// TIA Portal project "ağırlık" (V16)
// Vorlageprojekt für das Buch mit Zielsystem S7-1200

(* hardware
DEVICE "S7-1200-Station_1"  S7-1200 Station
   slot 0: "Baugruppenträger_0"  Rack  V1.0
   slot 1: "PLC_1"  CPU 1211C DC/DC/DC  6ES7 211-1AE40-0XB0  V4.1
DEVICE "HMI_1"  KTP700 Basic PN
   slot 0: "HMI_1"  KTP700 Basic PN  6AV2 123-2GB03-0AX0  16.0.0.0
   slot 1: "HMI_RT_1"  KTP700 Basic PN  6AV2 123-2GB03-0AX0  16.0.0.0
   slot 5: "HMI_1.IE_CP_1"  PROFINET Interface  16.0.0.0
      slot 1: "PROFINET Interface_1"  PROFINET Interface
         slot 1: "Port_1"  Port
*)

// ===== PLC "PLC_1"  CPU 1211C DC/DC/DC =====

VAR_GLOBAL   // PLC tag table "Default Table"
   "At scale entry" AT %I0.0 : Bool;
   "At scale" AT %I0.1 : Bool;
   "At scale exit" AT %I0.2 : Bool;
   "Left Pallet Sensor" AT %I0.3 : Bool;
   "At exit left" AT %I0.4 : Bool;
   "Front Palet sensor" AT %I0.5 : Bool;
   "At exit front" AT %I0.6 : Bool;
   "Right Pallet Sensor" AT %I0.7 : Bool;
   "At exit right" AT %I1.0 : Bool;
   "Start" AT %I1.1 : Bool;
   "Reset" AT %I1.2 : Bool;
   "Stop" AT %I1.3 : Bool;
   "FACTORY I/O (Running)" AT %I1.5 : Bool;
   "Pick & Place 1 (Box Detected)" AT %I1.6 : Bool;
   "Pick & Place 2 (Box Detected)" AT %I1.7 : Bool;
   "Pick & Place 3 (Box Detected)" AT %I2.0 : Bool;
   "Entry conveyor" AT %Q0.0 : Bool;
   "Load scale" AT %Q0.1 : Bool;
   "Send left" AT %Q0.2 : Bool;
   "Left conveyor" AT %Q0.3 : Bool;
   "Send right" AT %Q0.4 : Bool;
   "Right conveyor" AT %Q0.5 : Bool;
   "Send forward" AT %Q0.6 : Bool;
   "Front conveyor" AT %Q0.7 : Bool;
   "Start light" AT %Q1.0 : Bool;
   "Reset light" AT %Q1.1 : Bool;
   "Stop light" AT %Q1.2 : Bool;
   "Left Roller conveyor" AT %Q1.3 : Bool;
   "Right Roller Conveyor" AT %Q1.4 : Bool;
   "Front Roller conveyor" AT %Q1.5 : Bool;
END_VAR

VAR_GLOBAL   // PLC tag table "Tag table_1"
   "Pick & Place 1 X Position (V)" AT %ID34 : Real;
   "Pick & Place 1 Z Position (V)" AT %ID38 : Real;
   "Pick & Place 2 X Position (V)" AT %ID42 : Real;
   "Pick & Place 2 Z Position (V)" AT %ID46 : Real;
   "Pick & Place 3 X Position (V)" AT %ID50 : Real;
   "Pick & Place 3 Z Position (V)" AT %ID54 : Real;
   "Pick & Place 1 X Set Point (V)" AT %QD30 : Real;
   "Pick & Place 1 Y Set Point(V)" AT %QD34 : Real;
   "Pick & Place 1 Z Set Point (V)" AT %QD38 : Real;
   "Pick & Place 2 X Set Point (V)" AT %QD42 : Real;
   "Pick & Place 2 Z Set Point (V)" AT %QD46 : Real;
   "Pick & Place 3 X Set Point (V)" AT %QD50 : Real;
   "Pick & Place 3 Y Set Point(V)" AT %QD54 : Real;
   "Pick & Place 3 Z Set Point (V)" AT %QD58 : Real;
   "Weight" AT %ID30 : Real;
END_VAR

VAR_GLOBAL   // PLC tag table "Tag table_2"
   "tag1" AT %M0.0 : Bool;
   "tag2" AT %M0.1 : Bool;
   "tag3" AT %M0.2 : Bool;
   "Pick & Place 1 (Grab)" AT %Q1.7 : Bool;
   "Pick & Place 2 (Grab)" AT %Q2.1 : Bool;
   "Pick & Place 3 (Grab)" AT %Q2.3 : Bool;
END_VAR

DATA_BLOCK "Db"   // DB2
{ S7_Optimized_Access := 'TRUE' }
VERSION : 0.1
   VAR
      weight : Real;
      pallet_counter : Array[0..2] of DInt;
      "counter" : Array[0..3] of DInt;
      Weight_Value : Array[0..4] of Real;
      edge : Array[0..3] of Bool;
      palet_edge : Array[0..3] of Bool;
      hedef : DInt;
      hedef_percent : Real;
      doluluk_percent : Array[0..3] of Real;
      Total_count_normalized : Real;
      Doluluk_normalized : Array[0..3] of Real;
      Weight_Display : Real;
      Tartı_Hız : Time := T#1S;
      Pick_Place_Hız : Time := T#500MS;
      Total_Count : DInt;
      Start : Bool;
      Stop : Bool;
      Reset : Bool;
      Enable : Bool;
   END_VAR
BEGIN
   Weight_Value[0] := 2.5;
   Weight_Value[1] := 4.1;
   Weight_Value[2] := 4.5;
   Weight_Value[3] := 6.0;
   Weight_Value[4] := 7.0;
END_DATA_BLOCK

DATA_BLOCK "Pick_Place_DB"   // DB3
{ S7_Optimized_Access := 'TRUE' }
VERSION : 0.1
// stored: InstanceOfName Pick_Hafif
"Pick_Hafif"
BEGIN
END_DATA_BLOCK

DATA_BLOCK "Place_DB_4"   // DB8
{ S7_Optimized_Access := 'TRUE' }
VERSION : 0.1
// stored: InstanceOfName Place_Hafif
"Place_Hafif"
BEGIN
END_DATA_BLOCK

DATA_BLOCK "Place_DB_5"   // DB9
{ S7_Optimized_Access := 'TRUE' }
VERSION : 0.1
// stored: InstanceOfName Place_Hafif
"Place_Hafif"
BEGIN
END_DATA_BLOCK

DATA_BLOCK "Place_DB"   // DB10
{ S7_Optimized_Access := 'TRUE' }
VERSION : 0.1
// stored: InstanceOfName Place_Hafif
"Place_Hafif"
BEGIN
END_DATA_BLOCK

DATA_BLOCK "Place_DB_1"   // DB11
{ S7_Optimized_Access := 'TRUE' }
VERSION : 0.1
// stored: InstanceOfName Place_Hafif
"Place_Hafif"
BEGIN
END_DATA_BLOCK

DATA_BLOCK "Place_DB_2"   // DB12
{ S7_Optimized_Access := 'TRUE' }
VERSION : 0.1
// stored: InstanceOfName Place_Hafif
"Place_Hafif"
BEGIN
END_DATA_BLOCK

DATA_BLOCK "Place_DB_3"   // DB13
{ S7_Optimized_Access := 'TRUE' }
VERSION : 0.1
// stored: InstanceOfName Place_Hafif
"Place_Hafif"
BEGIN
END_DATA_BLOCK

DATA_BLOCK "Place_DB_6"   // DB14
{ S7_Optimized_Access := 'TRUE' }
VERSION : 0.1
// stored: InstanceOfName Place_Hafif
"Place_Hafif"
BEGIN
END_DATA_BLOCK

DATA_BLOCK "Place_DB_7"   // DB15
{ S7_Optimized_Access := 'TRUE' }
VERSION : 0.1
// stored: InstanceOfName Place_Hafif
"Place_Hafif"
BEGIN
END_DATA_BLOCK

DATA_BLOCK "Pick_Ağır_DB"   // DB16
{ S7_Optimized_Access := 'TRUE' }
VERSION : 0.1
// stored: InstanceOfName Pick_Ağır
"Pick_Ağır"
BEGIN
END_DATA_BLOCK

DATA_BLOCK "Pick_Orta_DB"   // DB17
{ S7_Optimized_Access := 'TRUE' }
VERSION : 0.1
// stored: InstanceOfName Pick_Orta
"Pick_Orta"
BEGIN
END_DATA_BLOCK

DATA_BLOCK "Place_Orta_DB"   // DB18
{ S7_Optimized_Access := 'TRUE' }
VERSION : 0.1
// stored: InstanceOfName Place_Orta
"Place_Orta"
BEGIN
END_DATA_BLOCK

DATA_BLOCK "Place_Ağır_DB"   // DB19
{ S7_Optimized_Access := 'TRUE' }
VERSION : 0.1
// stored: InstanceOfName Place_Ağır
"Place_Ağır"
BEGIN
END_DATA_BLOCK

// folder: System blocks/Program resources

DATA_BLOCK "IEC_Timer_0_DB_1"   // DB4
{ S7_Optimized_Access := 'TRUE' }
AUTHOR : Simatic
FAMILY : IEC
NAME : IEC_TMR
VERSION : 1.0
// stored: InstanceOfName IEC_TIMER
"IEC_TIMER"
BEGIN
END_DATA_BLOCK

DATA_BLOCK "IEC_Timer_0_DB"   // DB7
{ S7_Optimized_Access := 'TRUE' }
AUTHOR : Simatic
FAMILY : IEC
NAME : IEC_TMR
VERSION : 1.0
// stored: InstanceOfName IEC_TIMER
"IEC_TIMER"
BEGIN
END_DATA_BLOCK

DATA_BLOCK "IEC_Counter_0_DB_1"   // DB20
{ S7_Optimized_Access := 'TRUE' }
AUTHOR : Simatic
FAMILY : IEC
NAME : CNTR
VERSION : 1.0
// stored: InstanceOfName IEC_COUNTER
"IEC_COUNTER"
BEGIN
END_DATA_BLOCK

DATA_BLOCK "IEC_Counter_0_DB_2"   // DB22
{ S7_Optimized_Access := 'TRUE' }
AUTHOR : Simatic
FAMILY : IEC
NAME : CNTR
VERSION : 1.0
// stored: InstanceOfName IEC_COUNTER
"IEC_COUNTER"
BEGIN
END_DATA_BLOCK

DATA_BLOCK "IEC_Counter_0_DB_3"   // DB23
{ S7_Optimized_Access := 'TRUE' }
AUTHOR : Simatic
FAMILY : IEC
NAME : CNTR
VERSION : 1.0
// stored: InstanceOfName IEC_COUNTER
"IEC_COUNTER"
BEGIN
END_DATA_BLOCK

// folder: (top level)

FUNCTION_BLOCK "Pick_Hafif"   // FB1, LAD
{ S7_Optimized_Access := 'TRUE' }
VERSION : 0.1
   VAR
      state1 : Bool;
      state2 : Bool;
      IEC_Timer_0_Instance_3 : TON_TIME;
      IEC_Timer_0_Instance_4 : TON_TIME;
      IEC_Timer_0_Instance_5 : TON_TIME;
   END_VAR
BEGIN

REGION Network 1
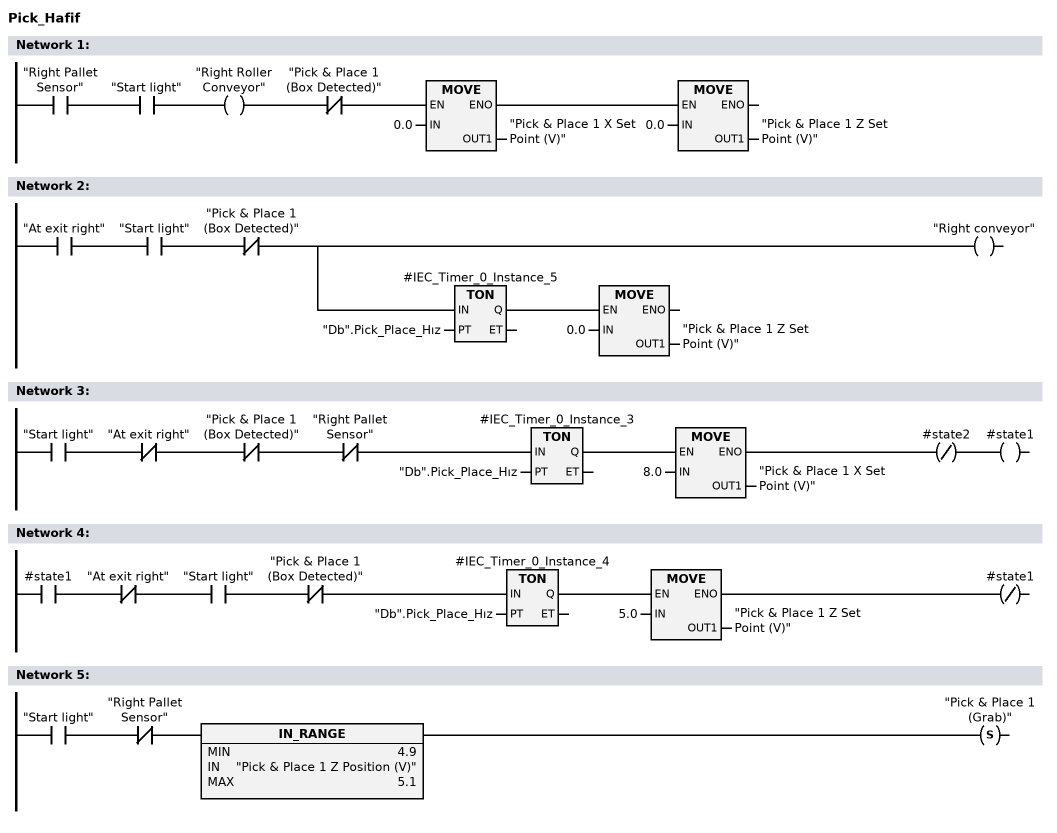
   "Right Roller Conveyor" := "Right Pallet Sensor" AND "Start light";
   IF "Right Roller Conveyor" AND NOT "Pick & Place 1 (Box Detected)" THEN
       "Pick & Place 1 X Set Point (V)" := 0.0;
       "Pick & Place 1 Z Set Point (V)" := 0.0;
   END_IF;
END_REGION

REGION Network 2
   "Right conveyor" := "At exit right" AND "Start light" AND NOT "Pick & Place 1 (Box Detected)";
   #IEC_Timer_0_Instance_5(IN := "Right conveyor", PT := "Db".Pick_Place_Hız);   // TON
   IF #IEC_Timer_0_Instance_5.Q THEN "Pick & Place 1 Z Set Point (V)" := 0.0; END_IF;
END_REGION

REGION Network 3
   #IEC_Timer_0_Instance_3(IN := "Start light" AND NOT "At exit right" AND NOT "Pick & Place 1 (Box Detected)" AND NOT "Right Pallet Sensor",   // TON
                           PT := "Db".Pick_Place_Hız);
   IF #IEC_Timer_0_Instance_3.Q THEN "Pick & Place 1 X Set Point (V)" := 8.0; END_IF;
   #state2 := NOT #IEC_Timer_0_Instance_3.Q;
   #state1 := #IEC_Timer_0_Instance_3.Q;
END_REGION

REGION Network 4
   #IEC_Timer_0_Instance_4(IN := #state1 AND NOT "At exit right" AND "Start light" AND NOT "Pick & Place 1 (Box Detected)",   // TON
                           PT := "Db".Pick_Place_Hız);
   IF #IEC_Timer_0_Instance_4.Q THEN "Pick & Place 1 Z Set Point (V)" := 5.0; END_IF;
   #state1 := NOT #IEC_Timer_0_Instance_4.Q;
END_REGION

REGION Network 5
   RUNG wire#powerrail
      Contact( "Start light" )
      I_Contact( "Right Pallet Sensor" )
      { S7_Templates := "SrcType := Real" } InRange(min := 4.9, in := "Pick & Place 1 Z Position (V)", max := 5.1)
      S_Coil( "Pick & Place 1 (Grab)" )
   END_RUNG
   // the same network as SCL:
   IF "Start light" AND NOT "Right Pallet Sensor" AND (4.9 <= "Pick & Place 1 Z Position (V)") AND ("Pick & Place 1 Z Position (V)" <= 5.1) THEN
       "Pick & Place 1 (Grab)" := TRUE;
   END_IF;
END_REGION
END_FUNCTION_BLOCK

FUNCTION_BLOCK "Place_Hafif"   // FB2, LAD
{ S7_Optimized_Access := 'TRUE' }
VERSION : 0.1
   VAR
      state1 : Bool;
      state2 : Bool;
      state3 : Bool;
      IEC_Timer_0_Instance_11 : TON_TIME;
      IEC_Timer_0_Instance_12 : TON_TIME;
      box : Int;
      IEC_Timer_0_Instance_13 : TON_TIME;
      R_TRIG_Instance : R_TRIG;
      edge : Bool;
      IEC_Timer_0_Instance_14 : TON_TIME;
      IEC_Timer_0_Instance_15 : TON_TIME;
      IEC_Timer_0_Instance_16 : TON_TIME;
   END_VAR
   VAR_TEMP   // added for the SCL form of the ladder/FBD networks
      _w1 : Bool;
   END_VAR
BEGIN

REGION Network 1
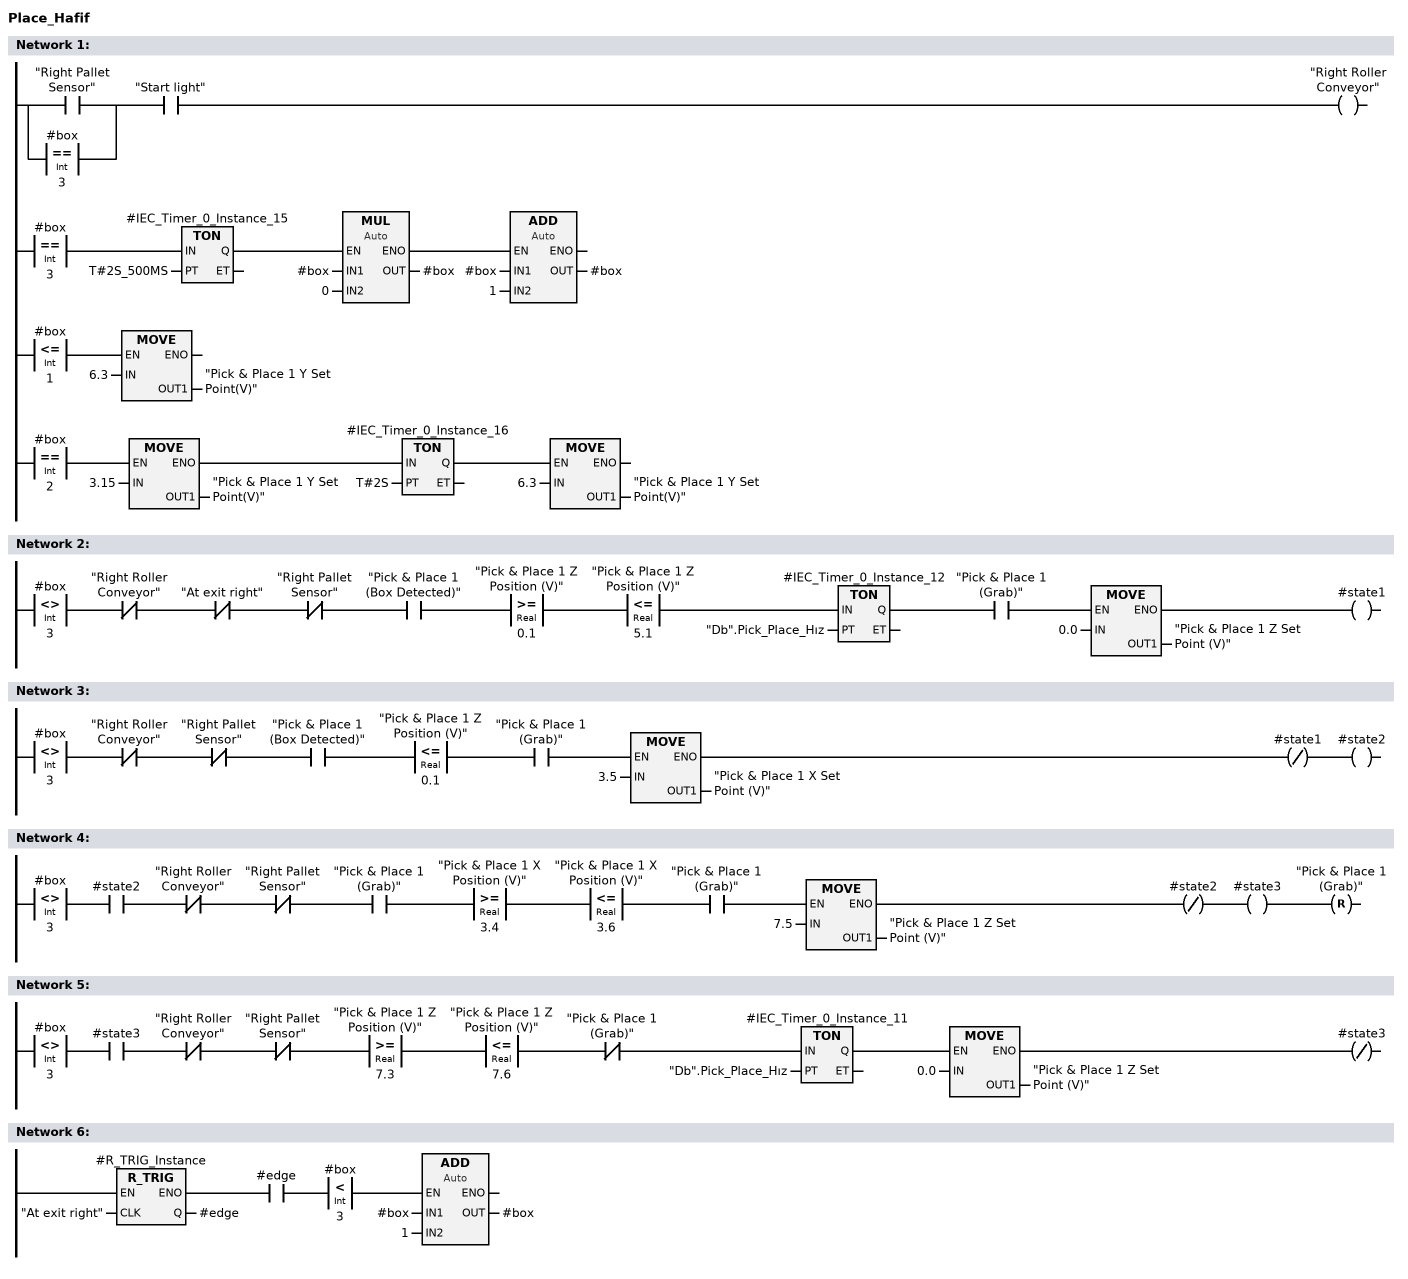
   "Right Roller Conveyor" := ("Right Pallet Sensor" OR (#box = 3)) AND "Start light";
   #IEC_Timer_0_Instance_15(IN := #box = 3, PT := T#2S_500MS);   // TON
   IF #IEC_Timer_0_Instance_15.Q THEN
       #box := #box * 0;
       #box := #box + 1;
   END_IF;
   IF #box <= 1 THEN "Pick & Place 1 Y Set Point(V)" := 6.3; END_IF;
   #_w1 := #box = 2;
   IF #_w1 THEN "Pick & Place 1 Y Set Point(V)" := 3.15; END_IF;
   #IEC_Timer_0_Instance_16(IN := #_w1, PT := T#2S);   // TON
   IF #IEC_Timer_0_Instance_16.Q THEN "Pick & Place 1 Y Set Point(V)" := 6.3; END_IF;
END_REGION

REGION Network 2
   #IEC_Timer_0_Instance_12(IN := (#box <> 3) AND NOT "Right Roller Conveyor" AND NOT "At exit right" AND NOT "Right Pallet Sensor" AND "Pick & Place 1 (Box Detected)" AND ("Pick & Place 1 Z Position (V)" >= 0.1) AND ("Pick & Place 1 Z Position (V)" <= 5.1),   // TON
                           PT := "Db".Pick_Place_Hız);
   #_w1 := #IEC_Timer_0_Instance_12.Q AND "Pick & Place 1 (Grab)";
   IF #_w1 THEN "Pick & Place 1 Z Set Point (V)" := 0.0; END_IF;
   #state1 := #_w1;
END_REGION

REGION Network 3
   #_w1 := (#box <> 3) AND NOT "Right Roller Conveyor" AND NOT "Right Pallet Sensor" AND "Pick & Place 1 (Box Detected)" AND ("Pick & Place 1 Z Position (V)" <= 0.1) AND "Pick & Place 1 (Grab)";
   IF #_w1 THEN "Pick & Place 1 X Set Point (V)" := 3.5; END_IF;
   #state1 := NOT #_w1;
   #state2 := #_w1;
END_REGION

REGION Network 4
   #_w1 := (#box <> 3) AND #state2 AND NOT "Right Roller Conveyor" AND NOT "Right Pallet Sensor" AND "Pick & Place 1 (Grab)" AND ("Pick & Place 1 X Position (V)" >= 3.4) AND ("Pick & Place 1 X Position (V)" <= 3.6) AND "Pick & Place 1 (Grab)";
   IF #_w1 THEN "Pick & Place 1 Z Set Point (V)" := 7.5; END_IF;
   #state2 := NOT #_w1;
   #state3 := #_w1;
   IF #_w1 THEN "Pick & Place 1 (Grab)" := FALSE; END_IF;
END_REGION

REGION Network 5
   #IEC_Timer_0_Instance_11(IN := (#box <> 3) AND #state3 AND NOT "Right Roller Conveyor" AND NOT "Right Pallet Sensor" AND ("Pick & Place 1 Z Position (V)" >= 7.3) AND ("Pick & Place 1 Z Position (V)" <= 7.6) AND NOT "Pick & Place 1 (Grab)",   // TON
                           PT := "Db".Pick_Place_Hız);
   IF #IEC_Timer_0_Instance_11.Q THEN "Pick & Place 1 Z Set Point (V)" := 0.0; END_IF;
   #state3 := NOT #IEC_Timer_0_Instance_11.Q;
END_REGION

REGION Network 6
   // ENO of a box is taken as its EN; it also drops when the box reports an error
   #R_TRIG_Instance(CLK := "At exit right", Q => #edge);   // R_TRIG
   IF #edge AND (#box < 3) THEN #box := #box + 1; END_IF;
END_REGION
END_FUNCTION_BLOCK

FUNCTION_BLOCK "Pick_Orta"   // FB3, LAD
{ S7_Optimized_Access := 'TRUE' }
VERSION : 0.1
   VAR
      state1 : Bool;
      state2 : Bool;
      IEC_Timer_0_Instance : TON_TIME;
      IEC_Timer_0_Instance_1 : TON_TIME;
      IEC_Timer_0_Instance_2 : TON_TIME;
   END_VAR
BEGIN

REGION Network 1
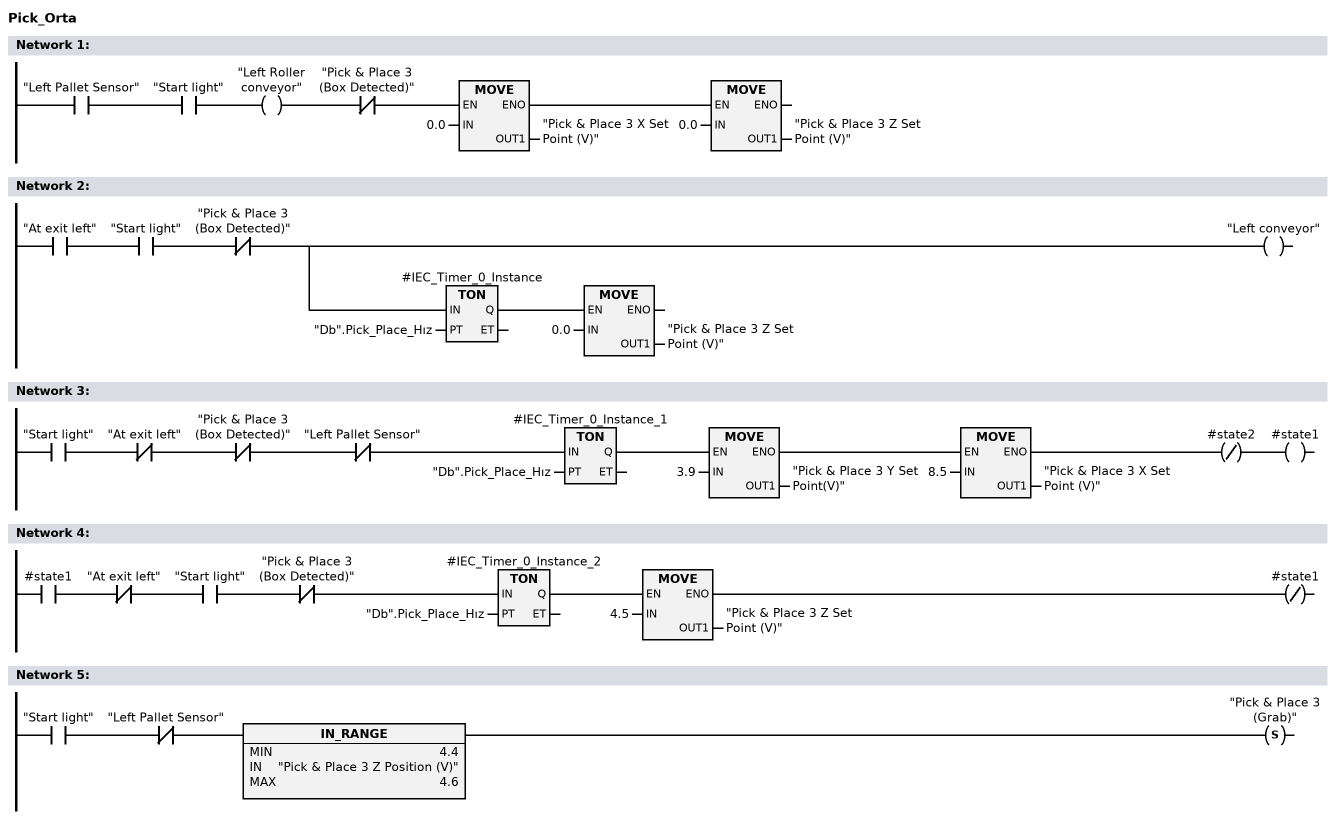
   "Left Roller conveyor" := "Left Pallet Sensor" AND "Start light";
   IF "Left Roller conveyor" AND NOT "Pick & Place 3 (Box Detected)" THEN
       "Pick & Place 3 X Set Point (V)" := 0.0;
       "Pick & Place 3 Z Set Point (V)" := 0.0;
   END_IF;
END_REGION

REGION Network 2
   "Left conveyor" := "At exit left" AND "Start light" AND NOT "Pick & Place 3 (Box Detected)";
   #IEC_Timer_0_Instance(IN := "Left conveyor", PT := "Db".Pick_Place_Hız);   // TON
   IF #IEC_Timer_0_Instance.Q THEN "Pick & Place 3 Z Set Point (V)" := 0.0; END_IF;
END_REGION

REGION Network 3
   #IEC_Timer_0_Instance_1(IN := "Start light" AND NOT "At exit left" AND NOT "Pick & Place 3 (Box Detected)" AND NOT "Left Pallet Sensor",   // TON
                           PT := "Db".Pick_Place_Hız);
   IF #IEC_Timer_0_Instance_1.Q THEN
       "Pick & Place 3 Y Set Point(V)" := 3.9;
       "Pick & Place 3 X Set Point (V)" := 8.5;
   END_IF;
   #state2 := NOT #IEC_Timer_0_Instance_1.Q;
   #state1 := #IEC_Timer_0_Instance_1.Q;
END_REGION

REGION Network 4
   #IEC_Timer_0_Instance_2(IN := #state1 AND NOT "At exit left" AND "Start light" AND NOT "Pick & Place 3 (Box Detected)",   // TON
                           PT := "Db".Pick_Place_Hız);
   IF #IEC_Timer_0_Instance_2.Q THEN "Pick & Place 3 Z Set Point (V)" := 4.5; END_IF;
   #state1 := NOT #IEC_Timer_0_Instance_2.Q;
END_REGION

REGION Network 5
   RUNG wire#powerrail
      Contact( "Start light" )
      I_Contact( "Left Pallet Sensor" )
      { S7_Templates := "SrcType := Real" } InRange(min := 4.4, in := "Pick & Place 3 Z Position (V)", max := 4.6)
      S_Coil( "Pick & Place 3 (Grab)" )
   END_RUNG
   // the same network as SCL:
   IF "Start light" AND NOT "Left Pallet Sensor" AND (4.4 <= "Pick & Place 3 Z Position (V)") AND ("Pick & Place 3 Z Position (V)" <= 4.6) THEN
       "Pick & Place 3 (Grab)" := TRUE;
   END_IF;
END_REGION
END_FUNCTION_BLOCK

FUNCTION_BLOCK "Place_Orta"   // FB4, LAD
{ S7_Optimized_Access := 'TRUE' }
VERSION : 0.1
   VAR
      state1 : Bool;
      state2 : Bool;
      state3 : Bool;
      edge : Bool;
      tag1 : Bool;
      box : Int;
      IEC_Timer_0_Instance_11 : TON_TIME;
      IEC_Timer_0_Instance_12 : TON_TIME;
      IEC_Timer_0_Instance : TON_TIME;
      IEC_Timer_0_Instance_1 : TON_TIME;
      R_TRIG_Instance : R_TRIG;
   END_VAR
   VAR_TEMP   // added for the SCL form of the ladder/FBD networks
      _w1 : Bool;
   END_VAR
BEGIN

REGION Network 1
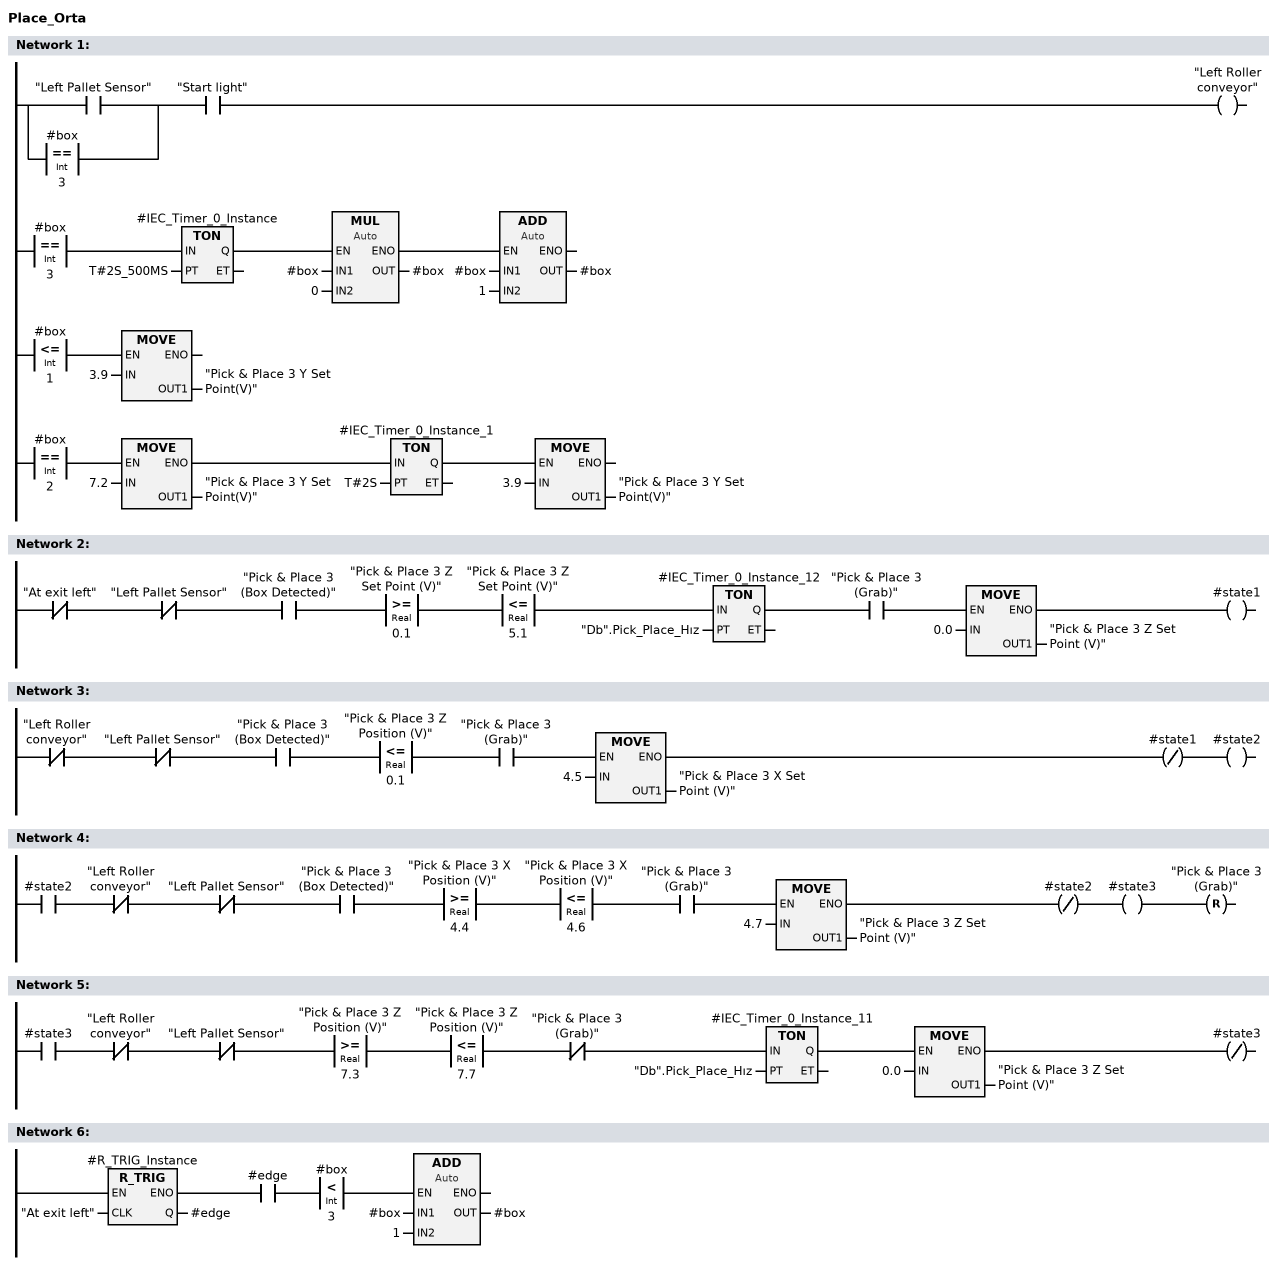
   "Left Roller conveyor" := ("Left Pallet Sensor" OR (#box = 3)) AND "Start light";
   #IEC_Timer_0_Instance(IN := #box = 3, PT := T#2S_500MS);   // TON
   IF #IEC_Timer_0_Instance.Q THEN
       #box := #box * 0;
       #box := #box + 1;
   END_IF;
   IF #box <= 1 THEN "Pick & Place 3 Y Set Point(V)" := 3.9; END_IF;
   #_w1 := #box = 2;
   IF #_w1 THEN "Pick & Place 3 Y Set Point(V)" := 7.2; END_IF;
   #IEC_Timer_0_Instance_1(IN := #_w1, PT := T#2S);   // TON
   IF #IEC_Timer_0_Instance_1.Q THEN "Pick & Place 3 Y Set Point(V)" := 3.9; END_IF;
END_REGION

REGION Network 2
   #IEC_Timer_0_Instance_12(IN := NOT "At exit left" AND NOT "Left Pallet Sensor" AND "Pick & Place 3 (Box Detected)" AND ("Pick & Place 3 Z Set Point (V)" >= 0.1) AND ("Pick & Place 3 Z Set Point (V)" <= 5.1),   // TON
                           PT := "Db".Pick_Place_Hız);
   #_w1 := #IEC_Timer_0_Instance_12.Q AND "Pick & Place 3 (Grab)";
   IF #_w1 THEN "Pick & Place 3 Z Set Point (V)" := 0.0; END_IF;
   #state1 := #_w1;
END_REGION

REGION Network 3
   #_w1 := NOT "Left Roller conveyor" AND NOT "Left Pallet Sensor" AND "Pick & Place 3 (Box Detected)" AND ("Pick & Place 3 Z Position (V)" <= 0.1) AND "Pick & Place 3 (Grab)";
   IF #_w1 THEN "Pick & Place 3 X Set Point (V)" := 4.5; END_IF;
   #state1 := NOT #_w1;
   #state2 := #_w1;
END_REGION

REGION Network 4
   #_w1 := #state2 AND NOT "Left Roller conveyor" AND NOT "Left Pallet Sensor" AND "Pick & Place 3 (Box Detected)" AND ("Pick & Place 3 X Position (V)" >= 4.4) AND ("Pick & Place 3 X Position (V)" <= 4.6) AND "Pick & Place 3 (Grab)";
   IF #_w1 THEN "Pick & Place 3 Z Set Point (V)" := 4.7; END_IF;
   #state2 := NOT #_w1;
   #state3 := #_w1;
   IF #_w1 THEN "Pick & Place 3 (Grab)" := FALSE; END_IF;
END_REGION

REGION Network 5
   #IEC_Timer_0_Instance_11(IN := #state3 AND NOT "Left Roller conveyor" AND NOT "Left Pallet Sensor" AND ("Pick & Place 3 Z Position (V)" >= 7.3) AND ("Pick & Place 3 Z Position (V)" <= 7.7) AND NOT "Pick & Place 3 (Grab)",   // TON
                           PT := "Db".Pick_Place_Hız);
   IF #IEC_Timer_0_Instance_11.Q THEN "Pick & Place 3 Z Set Point (V)" := 0.0; END_IF;
   #state3 := NOT #IEC_Timer_0_Instance_11.Q;
END_REGION

REGION Network 6
   // ENO of a box is taken as its EN; it also drops when the box reports an error
   #R_TRIG_Instance(CLK := "At exit left", Q => #edge);   // R_TRIG
   IF #edge AND (#box < 3) THEN #box := #box + 1; END_IF;
END_REGION
END_FUNCTION_BLOCK

FUNCTION_BLOCK "Pick_Ağır"   // FB5, LAD
{ S7_Optimized_Access := 'TRUE' }
VERSION : 0.1
   VAR
      state1 : Bool;
      state2 : Bool;
      state3 : Bool;
      IEC_Timer_0_Instance : TON_TIME;
      IEC_Timer_0_Instance_1 : TON_TIME;
      IEC_Timer_0_Instance_2 : TON_TIME;
   END_VAR
   VAR_TEMP   // added for the SCL form of the ladder/FBD networks
      _w1 : Bool;
   END_VAR
BEGIN

REGION Network 1
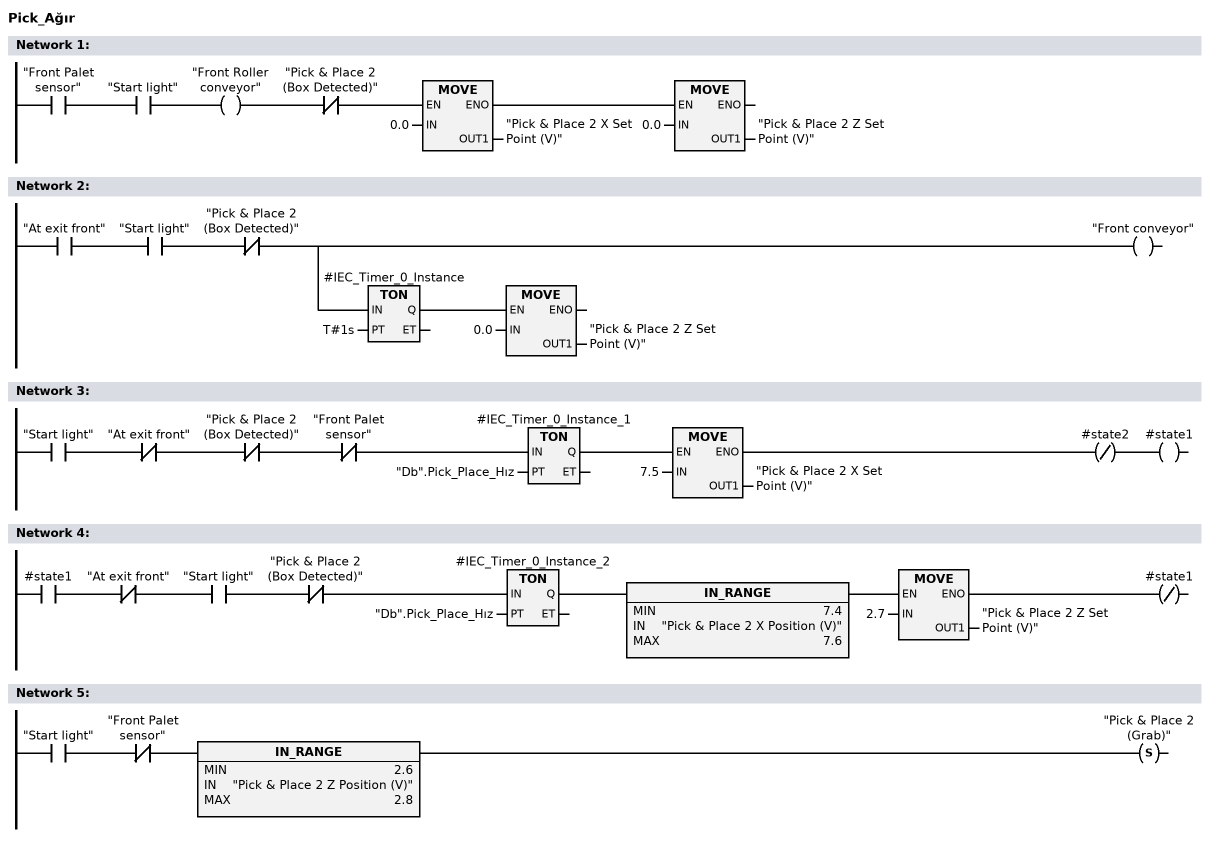
   "Front Roller conveyor" := "Front Palet sensor" AND "Start light";
   IF "Front Roller conveyor" AND NOT "Pick & Place 2 (Box Detected)" THEN
       "Pick & Place 2 X Set Point (V)" := 0.0;
       "Pick & Place 2 Z Set Point (V)" := 0.0;
   END_IF;
END_REGION

REGION Network 2
   "Front conveyor" := "At exit front" AND "Start light" AND NOT "Pick & Place 2 (Box Detected)";
   #IEC_Timer_0_Instance(IN := "Front conveyor", PT := T#1s);   // TON
   IF #IEC_Timer_0_Instance.Q THEN "Pick & Place 2 Z Set Point (V)" := 0.0; END_IF;
END_REGION

REGION Network 3
   #IEC_Timer_0_Instance_1(IN := "Start light" AND NOT "At exit front" AND NOT "Pick & Place 2 (Box Detected)" AND NOT "Front Palet sensor",   // TON
                           PT := "Db".Pick_Place_Hız);
   IF #IEC_Timer_0_Instance_1.Q THEN "Pick & Place 2 X Set Point (V)" := 7.5; END_IF;
   #state2 := NOT #IEC_Timer_0_Instance_1.Q;
   #state1 := #IEC_Timer_0_Instance_1.Q;
END_REGION

REGION Network 4
   #IEC_Timer_0_Instance_2(IN := #state1 AND NOT "At exit front" AND "Start light" AND NOT "Pick & Place 2 (Box Detected)",   // TON
                           PT := "Db".Pick_Place_Hız);
   #_w1 := #IEC_Timer_0_Instance_2.Q AND (7.4 <= "Pick & Place 2 X Position (V)") AND ("Pick & Place 2 X Position (V)" <= 7.6);
   IF #_w1 THEN "Pick & Place 2 Z Set Point (V)" := 2.7; END_IF;
   #state1 := NOT #_w1;
END_REGION

REGION Network 5
   RUNG wire#powerrail
      Contact( "Start light" )
      I_Contact( "Front Palet sensor" )
      { S7_Templates := "SrcType := Real" } InRange(min := 2.6, in := "Pick & Place 2 Z Position (V)", max := 2.8)
      S_Coil( "Pick & Place 2 (Grab)" )
   END_RUNG
   // the same network as SCL:
   IF "Start light" AND NOT "Front Palet sensor" AND (2.6 <= "Pick & Place 2 Z Position (V)") AND ("Pick & Place 2 Z Position (V)" <= 2.8) THEN
       "Pick & Place 2 (Grab)" := TRUE;
   END_IF;
END_REGION
END_FUNCTION_BLOCK

FUNCTION_BLOCK "Place_Ağır"   // FB6, LAD
{ S7_Optimized_Access := 'TRUE' }
VERSION : 0.1
   VAR
      IEC_Timer_0_Instance : TON_TIME;
      IEC_Timer_0_Instance_1 : TON_TIME;
      state1 : Bool;
      state2 : Bool;
      state3 : Bool;
      edge : Bool;
      box : Int;
      R_TRIG_Instance : R_TRIG;
   END_VAR
   VAR_TEMP   // added for the SCL form of the ladder/FBD networks
      _w1 : Bool;
   END_VAR
BEGIN

REGION Network 1
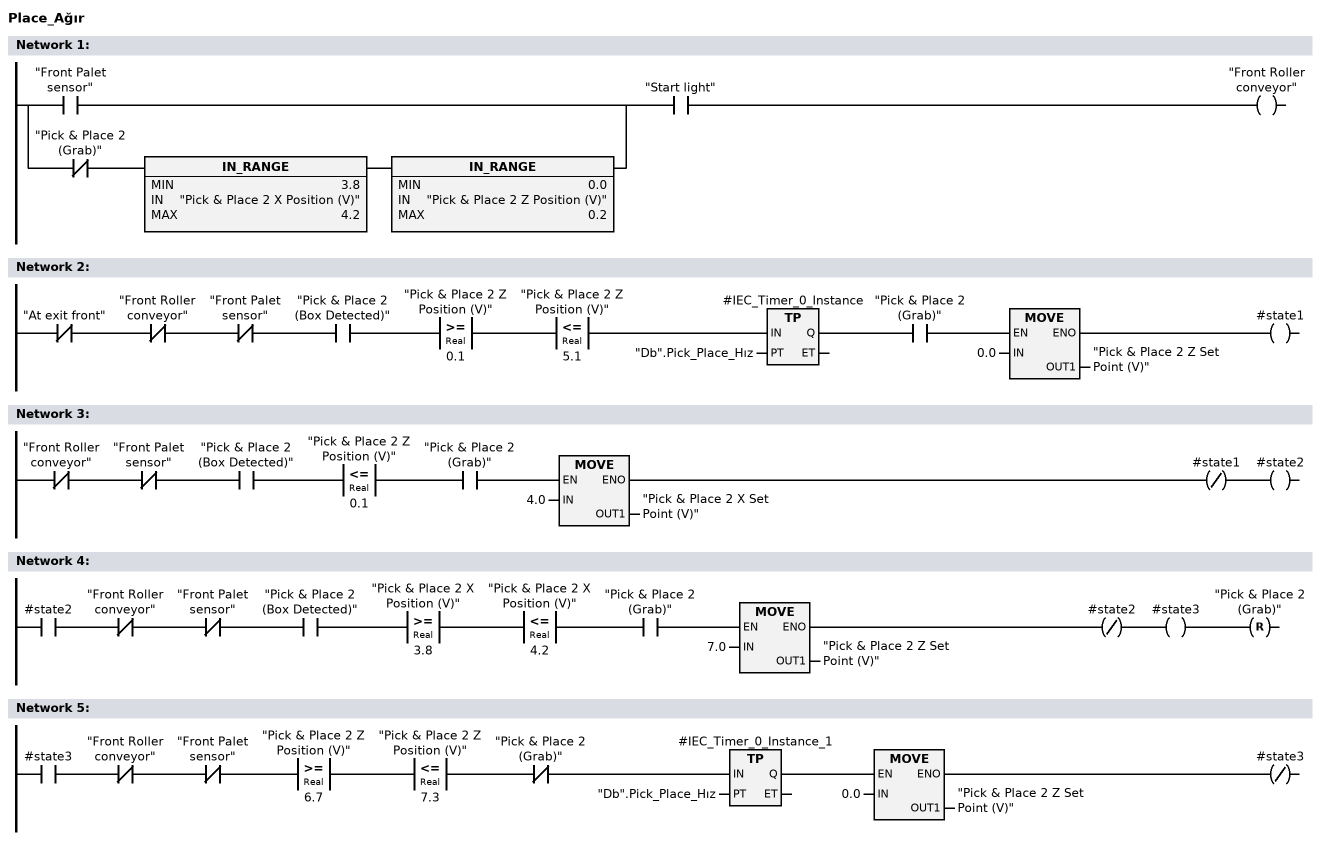
   RUNG wire#powerrail
      Contact( "Front Palet sensor" )
      wire#w1
      Contact( "Start light" )
      Coil( "Front Roller conveyor" )
   END_RUNG
   RUNG wire#powerrail
      I_Contact( "Pick & Place 2 (Grab)" )
      { S7_Templates := "SrcType := Real" } InRange(min := 3.8, in := "Pick & Place 2 X Position (V)", max := 4.2)
      { S7_Templates := "SrcType := Real" } InRange(min := 0.0, in := "Pick & Place 2 Z Position (V)", max := 0.2)
   END_RUNG wire#w1
   // the same network as SCL:
   "Front Roller conveyor" := ("Front Palet sensor" OR (NOT "Pick & Place 2 (Grab)" AND (3.8 <= "Pick & Place 2 X Position (V)") AND ("Pick & Place 2 X Position (V)" <= 4.2) AND (0.0 <= "Pick & Place 2 Z Position (V)") AND ("Pick & Place 2 Z Position (V)" <= 0.2))) AND "Start light";
END_REGION

REGION Network 2
   #IEC_Timer_0_Instance(IN := NOT "At exit front" AND NOT "Front Roller conveyor" AND NOT "Front Palet sensor" AND "Pick & Place 2 (Box Detected)" AND ("Pick & Place 2 Z Position (V)" >= 0.1) AND ("Pick & Place 2 Z Position (V)" <= 5.1),   // TP
                         PT := "Db".Pick_Place_Hız);
   #_w1 := #IEC_Timer_0_Instance.Q AND "Pick & Place 2 (Grab)";
   IF #_w1 THEN "Pick & Place 2 Z Set Point (V)" := 0.0; END_IF;
   #state1 := #_w1;
END_REGION

REGION Network 3
   #_w1 := NOT "Front Roller conveyor" AND NOT "Front Palet sensor" AND "Pick & Place 2 (Box Detected)" AND ("Pick & Place 2 Z Position (V)" <= 0.1) AND "Pick & Place 2 (Grab)";
   IF #_w1 THEN "Pick & Place 2 X Set Point (V)" := 4.0; END_IF;
   #state1 := NOT #_w1;
   #state2 := #_w1;
END_REGION

REGION Network 4
   #_w1 := #state2 AND NOT "Front Roller conveyor" AND NOT "Front Palet sensor" AND "Pick & Place 2 (Box Detected)" AND ("Pick & Place 2 X Position (V)" >= 3.8) AND ("Pick & Place 2 X Position (V)" <= 4.2) AND "Pick & Place 2 (Grab)";
   IF #_w1 THEN "Pick & Place 2 Z Set Point (V)" := 7.0; END_IF;
   #state2 := NOT #_w1;
   #state3 := #_w1;
   IF #_w1 THEN "Pick & Place 2 (Grab)" := FALSE; END_IF;
END_REGION

REGION Network 5
   #IEC_Timer_0_Instance_1(IN := #state3 AND NOT "Front Roller conveyor" AND NOT "Front Palet sensor" AND ("Pick & Place 2 Z Position (V)" >= 6.7) AND ("Pick & Place 2 Z Position (V)" <= 7.3) AND NOT "Pick & Place 2 (Grab)",   // TP
                           PT := "Db".Pick_Place_Hız);
   IF #IEC_Timer_0_Instance_1.Q THEN "Pick & Place 2 Z Set Point (V)" := 0.0; END_IF;
   #state3 := NOT #IEC_Timer_0_Instance_1.Q;
END_REGION
END_FUNCTION_BLOCK

FUNCTION "Tartı" : Void   // FC1, LAD
{ S7_Optimized_Access := 'TRUE' }
VERSION : 0.1
   VAR_INPUT
      at_scale_entry_sensor : Bool;
      start_light : Bool;
      at_scale_sensor : Bool;
      weight_display : Real;
   END_VAR
   VAR_OUTPUT
      "right roller" : Bool;
      "left roller" : Bool;
      "front roller" : Bool;
      load_scale : Bool;
      entry_conveyor : Bool;
   END_VAR
   VAR_TEMP   // added for the SCL form of the ladder/FBD networks
      _w1 : Bool;
   END_VAR
BEGIN

REGION Network 1
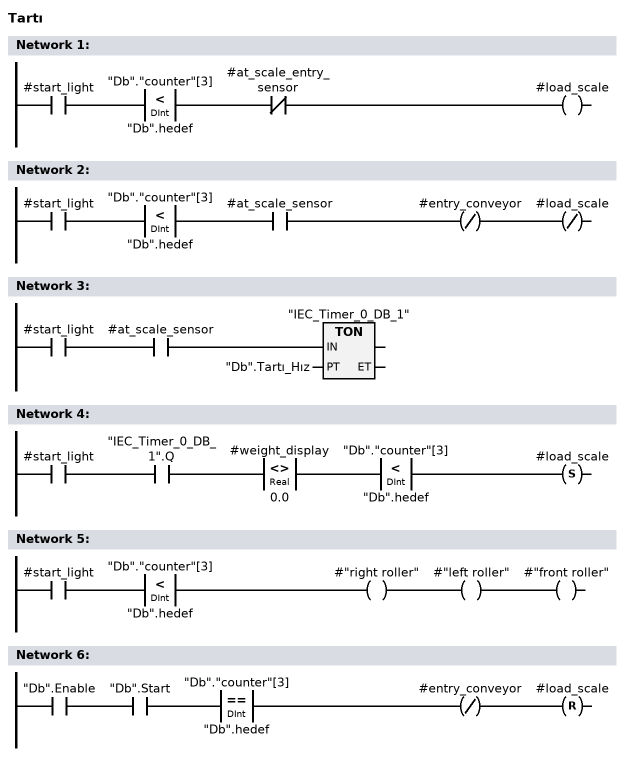
   RUNG wire#powerrail
      Contact( #start_light )
      { S7_Templates := "SrcType := DInt" } LT_Contact(in1 := "Db"."counter"[3], in2 := "Db".hedef)
      I_Contact( #at_scale_entry_sensor )
      Coil( #load_scale )
   END_RUNG
   // the same network as SCL:
   #load_scale := #start_light AND ("Db"."counter"[3] < "Db".hedef) AND NOT #at_scale_entry_sensor;
END_REGION

REGION Network 2
   RUNG wire#powerrail
      Contact( #start_light )
      { S7_Templates := "SrcType := DInt" } LT_Contact(in1 := "Db"."counter"[3], in2 := "Db".hedef)
      Contact( #at_scale_sensor )
      I_Coil( #entry_conveyor )
      I_Coil( #load_scale )
   END_RUNG
   // the same network as SCL:
   #_w1 := #start_light AND ("Db"."counter"[3] < "Db".hedef) AND #at_scale_sensor;
   #entry_conveyor := NOT #_w1;
   #load_scale := NOT #_w1;
END_REGION

REGION Network 3
   "IEC_Timer_0_DB_1".TON(IN := #start_light AND #at_scale_sensor, PT := "Db".Tartı_Hız);
END_REGION

REGION Network 4
   RUNG wire#powerrail
      Contact( #start_light )
      Contact( "IEC_Timer_0_DB_1".Q )
      { S7_Templates := "SrcType := Real" } NE_Contact(in1 := #weight_display, in2 := 0.0)
      { S7_Templates := "SrcType := DInt" } LT_Contact(in1 := "Db"."counter"[3], in2 := "Db".hedef)
      S_Coil( #load_scale )
   END_RUNG
   // the same network as SCL:
   IF #start_light AND "IEC_Timer_0_DB_1".Q AND (#weight_display <> 0.0) AND ("Db"."counter"[3] < "Db".hedef) THEN
       #load_scale := TRUE;
   END_IF;
END_REGION

REGION Network 5
   RUNG wire#powerrail
      Contact( #start_light )
      { S7_Templates := "SrcType := DInt" } LT_Contact(in1 := "Db"."counter"[3], in2 := "Db".hedef)
      Coil( #"right roller" )
      Coil( #"left roller" )
      Coil( #"front roller" )
   END_RUNG
   // the same network as SCL:
   #"right roller" := #start_light AND ("Db"."counter"[3] < "Db".hedef);
   #"left roller" := #"right roller";
   #"front roller" := #"right roller";
END_REGION

REGION Network 6
   RUNG wire#powerrail
      Contact( "Db".Enable )
      Contact( "Db".Start )
      { S7_Templates := "SrcType := DInt" } EQ_Contact(in1 := "Db"."counter"[3], in2 := "Db".hedef)
      I_Coil( #entry_conveyor )
      R_Coil( #load_scale )
   END_RUNG
   // the same network as SCL:
   #_w1 := "Db".Enable AND "Db".Start AND ("Db"."counter"[3] = "Db".hedef);
   #entry_conveyor := NOT #_w1;
   IF #_w1 THEN #load_scale := FALSE; END_IF;
END_REGION
END_FUNCTION

FUNCTION "Sınıflandırma" : Void   // FC2, LAD
{ S7_Optimized_Access := 'TRUE' }
VERSION : 0.1
   VAR_INPUT
      weight_display : Real;
      enable : Bool;
      hedef : DInt;
      right_sensor : Bool;
      left_sensor : Bool;
      forward_sensor : Bool;
      weight : Array[0..4] of Real;
   END_VAR
   VAR_OUTPUT
      forward : Bool;
      right : Bool;
      left : Bool;
   END_VAR
   VAR_IN_OUT
      counter1 : DInt;
      counter2 : DInt;
      counter3 : DInt;
      counter4 : DInt;
   END_VAR
   VAR_TEMP   // added for the SCL form of the ladder/FBD networks
      _w1 : Bool;
   END_VAR
BEGIN

REGION Network 1
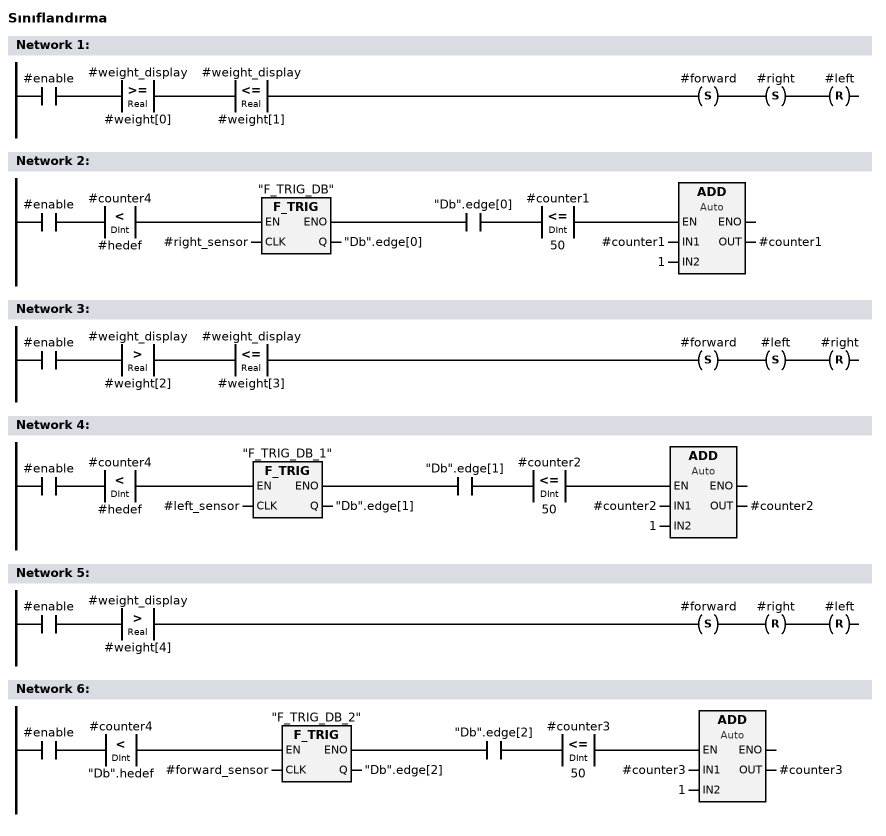
   RUNG wire#powerrail
      Contact( #enable )
      { S7_Templates := "SrcType := Real" } GE_Contact(in1 := #weight_display, in2 := #weight[0])
      { S7_Templates := "SrcType := Real" } LE_Contact(in1 := #weight_display, in2 := #weight[1])
      S_Coil( #forward )
      S_Coil( #right )
      R_Coil( #left )
   END_RUNG
   // the same network as SCL:
   IF #enable AND (#weight_display >= #weight[0]) AND (#weight_display <= #weight[1]) THEN
       #forward := TRUE;
       #right := TRUE;
       #left := FALSE;
   END_IF;
END_REGION

REGION Network 2
   // ENO of a box is taken as its EN; it also drops when the box reports an error
   #_w1 := #enable AND (#counter4 < #hedef);
   IF #_w1 THEN
       "F_TRIG_DB"(CLK := #right_sensor, Q => "Db".edge[0]);   // F_TRIG
   END_IF;
   IF #_w1 AND "Db".edge[0] AND (#counter1 <= 50) THEN #counter1 := #counter1 + 1; END_IF;
END_REGION

REGION Network 3
   RUNG wire#powerrail
      Contact( #enable )
      { S7_Templates := "SrcType := Real" } GT_Contact(in1 := #weight_display, in2 := #weight[2])
      { S7_Templates := "SrcType := Real" } LE_Contact(in1 := #weight_display, in2 := #weight[3])
      S_Coil( #forward )
      S_Coil( #left )
      R_Coil( #right )
   END_RUNG
   // the same network as SCL:
   IF #enable AND (#weight_display > #weight[2]) AND (#weight_display <= #weight[3]) THEN
       #forward := TRUE;
       #left := TRUE;
       #right := FALSE;
   END_IF;
END_REGION

REGION Network 4
   // ENO of a box is taken as its EN; it also drops when the box reports an error
   #_w1 := #enable AND (#counter4 < #hedef);
   IF #_w1 THEN
       "F_TRIG_DB_1"(CLK := #left_sensor, Q => "Db".edge[1]);   // F_TRIG
   END_IF;
   IF #_w1 AND "Db".edge[1] AND (#counter2 <= 50) THEN #counter2 := #counter2 + 1; END_IF;
END_REGION

REGION Network 5
   RUNG wire#powerrail
      Contact( #enable )
      { S7_Templates := "SrcType := Real" } GT_Contact(in1 := #weight_display, in2 := #weight[4])
      S_Coil( #forward )
      R_Coil( #right )
      R_Coil( #left )
   END_RUNG
   // the same network as SCL:
   IF #enable AND (#weight_display > #weight[4]) THEN
       #forward := TRUE;
       #right := FALSE;
       #left := FALSE;
   END_IF;
END_REGION

REGION Network 6
   // ENO of a box is taken as its EN; it also drops when the box reports an error
   #_w1 := #enable AND (#counter4 < "Db".hedef);
   IF #_w1 THEN
       "F_TRIG_DB_2"(CLK := #forward_sensor, Q => "Db".edge[2]);   // F_TRIG
   END_IF;
   IF #_w1 AND "Db".edge[2] AND (#counter3 <= 50) THEN #counter3 := #counter3 + 1; END_IF;
END_REGION
END_FUNCTION

FUNCTION "MHJ-PLC-Lab-Function-S71200" : Void   // FC9000, SCL
{ S7_Optimized_Access := 'TRUE' }
VERSION : 0.1
   VAR_TEMP
      rdTimeReturn : Int;
      outputTime : DTL;
      SyncVal : Byte;
      forVal : Int;
      forVal_2 : Int;
      Value : Byte;
   END_VAR
   VAR CONSTANT
      CompVal : Byte := 16#34;
      Value_01 : Byte := 16#11;
      Value_01_DW : DWord := 16#A165_D992;
      Value_02_DW : DWord := 16#58BE_4401;
   END_VAR
BEGIN

   #Value:=PEEK(area := 16#82,
        dbNumber := 0,
        byteOffset := 511);
   #Value := #Value + 1;

   POKE(area := 16#82,
        dbNumber := 0,
        byteOffset := 511,
        value := #Value);

   POKE(area:=16#81,
        dbNumber:=0,
        byteOffset:=1016,
        value:=#Value_01_DW);
   POKE(area := 16#81,
        dbNumber := 0,
        byteOffset := 1020,
        value := #Value_02_DW);

   POKE(area := 16#81,
        dbNumber := 0,
        byteOffset := 511,
        value := B#16#00);

   FOR #forVal := 0 TO 120 DO
       FOR #forVal_2:=0 TO 10 DO
           #rdTimeReturn:=RD_SYS_T(#outputTime);
           #rdTimeReturn := WR_SYS_T(#outputTime);
           #rdTimeReturn := RD_SYS_T(#outputTime);
           #rdTimeReturn := WR_SYS_T(#outputTime);
       END_FOR;
       #SyncVal:= PEEK(area := 16#81,
                      dbNumber := 0,
                      byteOffset := 511);
       IF #SyncVal = #CompVal THEN
          GOTO M_1;
       END_IF;
   END_FOR;
   RETURN;

   M_1:
   POKE(area := 16#81,
        dbNumber := 0,
        byteOffset := 511,
        value := B#16#0);
END_FUNCTION

ORGANIZATION_BLOCK "Main"   // OB1, LAD, ProgramCycle
TITLE = "Main Program Sweep (Cycle)"
{ S7_Optimized_Access := 'TRUE' }
VERSION : 0.1
   VAR_INPUT
      Initial_Call : Bool;   // Initial call of this OB
      Remanence : Bool;   // =True, if remanent data are available
   END_VAR
   VAR_TEMP   // added for the SCL form of the ladder/FBD networks
      _w1 : Bool;
   END_VAR
BEGIN

REGION Network 1
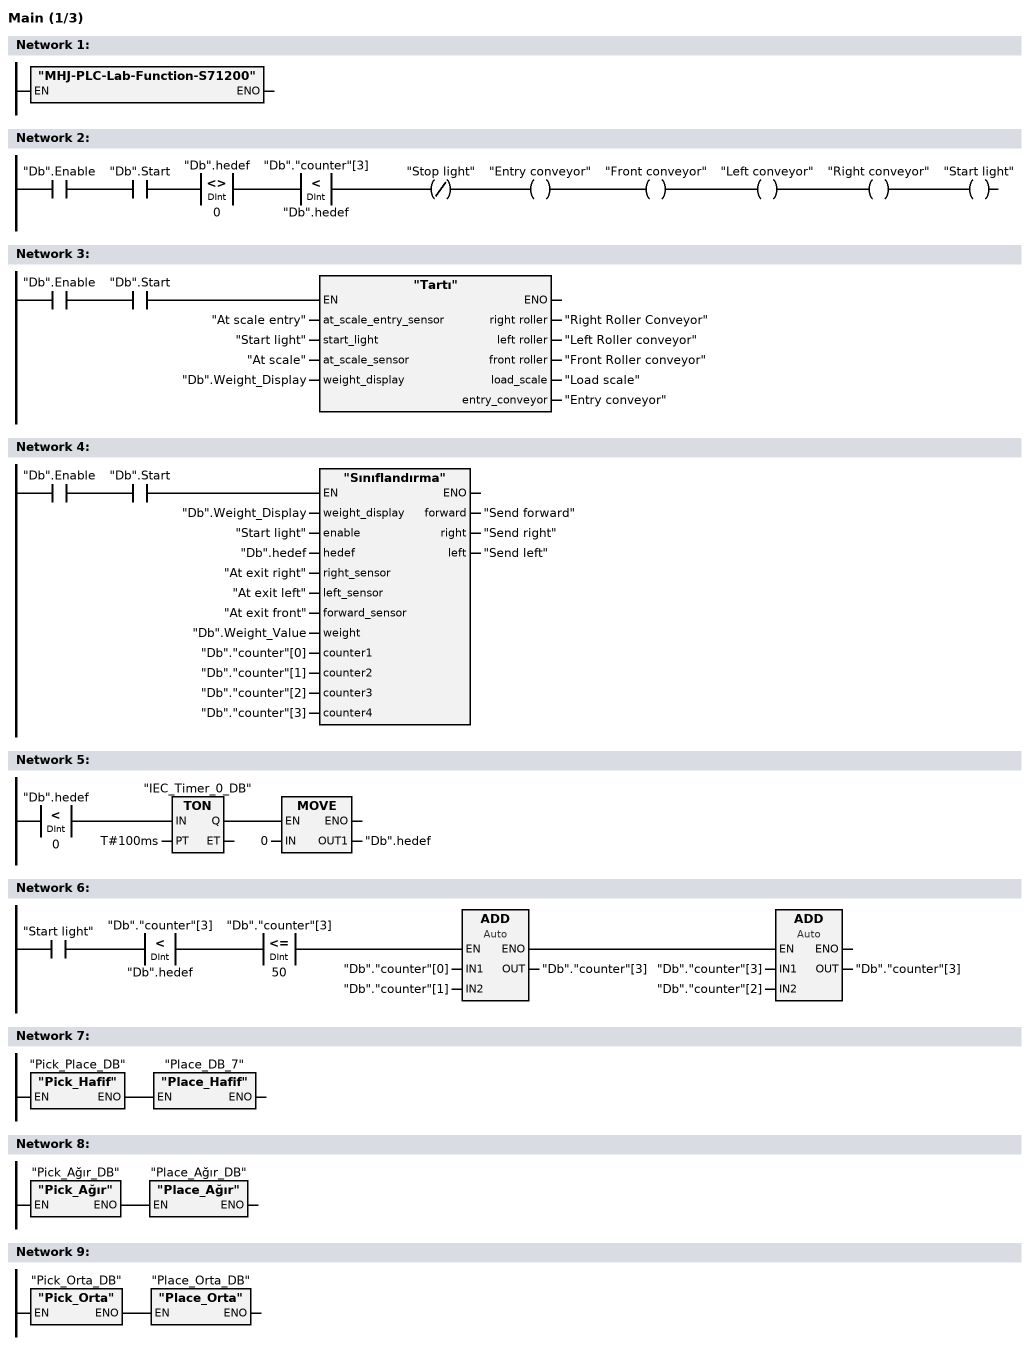
   RUNG wire#powerrail
      "MHJ-PLC-Lab-Function-S71200"()
   END_RUNG
   // the same network as SCL:
   "MHJ-PLC-Lab-Function-S71200"();
END_REGION

REGION Network 2
   RUNG wire#powerrail
      Contact( "Db".Enable )
      Contact( "Db".Start )
      { S7_Templates := "SrcType := DInt" } NE_Contact(in1 := "Db".hedef, in2 := 0)
      { S7_Templates := "SrcType := DInt" } LT_Contact(in1 := "Db"."counter"[3], in2 := "Db".hedef)
      I_Coil( "Stop light" )
      Coil( "Entry conveyor" )
      Coil( "Front conveyor" )
      Coil( "Left conveyor" )
      Coil( "Right conveyor" )
      Coil( "Start light" )
   END_RUNG
   // the same network as SCL:
   #_w1 := "Db".Enable AND "Db".Start AND ("Db".hedef <> 0) AND ("Db"."counter"[3] < "Db".hedef);
   "Stop light" := NOT #_w1;
   "Entry conveyor" := #_w1;
   "Front conveyor" := #_w1;
   "Left conveyor" := #_w1;
   "Right conveyor" := #_w1;
   "Start light" := #_w1;
END_REGION

REGION Network 3
   RUNG wire#powerrail
      Contact( "Db".Enable )
      Contact( "Db".Start )
      "Tartı"(at_scale_entry_sensor := "At scale entry", start_light := "Start light", at_scale_sensor := "At scale", weight_display := "Db".Weight_Display, "right roller" => "Right Roller Conveyor", "left roller" => "Left Roller conveyor", "front roller" => "Front Roller conveyor", load_scale => "Load scale", entry_conveyor => "Entry conveyor")
   END_RUNG
   // the same network as SCL:
   IF "Db".Enable AND "Db".Start THEN
       "Tartı"(at_scale_entry_sensor := "At scale entry",
               start_light := "Start light",
               at_scale_sensor := "At scale",
               weight_display := "Db".Weight_Display,
               "right roller" => "Right Roller Conveyor",
               "left roller" => "Left Roller conveyor",
               "front roller" => "Front Roller conveyor",
               load_scale => "Load scale",
               entry_conveyor => "Entry conveyor");
   END_IF;
END_REGION

REGION Network 4
   RUNG wire#powerrail
      Contact( "Db".Enable )
      Contact( "Db".Start )
      "Sınıflandırma"(weight_display := "Db".Weight_Display, enable := "Start light", hedef := "Db".hedef, right_sensor := "At exit right", left_sensor := "At exit left", forward_sensor := "At exit front", weight := "Db".Weight_Value, counter1 := "Db"."counter"[0], counter2 := "Db"."counter"[1], counter3 := "Db"."counter"[2], counter4 := "Db"."counter"[3], forward => "Send forward", right => "Send right", left => "Send left")
   END_RUNG
   // the same network as SCL:
   IF "Db".Enable AND "Db".Start THEN
       "Sınıflandırma"(weight_display := "Db".Weight_Display,
                       enable := "Start light",
                       hedef := "Db".hedef,
                       right_sensor := "At exit right",
                       left_sensor := "At exit left",
                       forward_sensor := "At exit front",
                       weight := "Db".Weight_Value,
                       counter1 := "Db"."counter"[0],
                       counter2 := "Db"."counter"[1],
                       counter3 := "Db"."counter"[2],
                       counter4 := "Db"."counter"[3],
                       forward => "Send forward",
                       right => "Send right",
                       left => "Send left");
   END_IF;
END_REGION

REGION Network 5
   "IEC_Timer_0_DB".TON(IN := "Db".hedef < 0, PT := T#100ms);
   IF "IEC_Timer_0_DB".Q THEN "Db".hedef := 0; END_IF;
END_REGION

REGION Network 6
   RUNG wire#powerrail
      Contact( "Start light" )
      { S7_Templates := "SrcType := DInt" } LT_Contact(in1 := "Db"."counter"[3], in2 := "Db".hedef)
      { S7_Templates := "SrcType := DInt" } LE_Contact(in1 := "Db"."counter"[3], in2 := 50)
      Add(in1 := "Db"."counter"[0], in2 := "Db"."counter"[1], out => "Db"."counter"[3])
      Add(in1 := "Db"."counter"[3], in2 := "Db"."counter"[2], out => "Db"."counter"[3])
   END_RUNG
   // the same network as SCL:
   #_w1 := "Start light" AND ("Db"."counter"[3] < "Db".hedef) AND ("Db"."counter"[3] <= 50);
   IF #_w1 THEN
       "Db"."counter"[3] := "Db"."counter"[0] + "Db"."counter"[1];
       "Db"."counter"[3] := "Db"."counter"[3] + "Db"."counter"[2];
   END_IF;
END_REGION

REGION Network 7
   RUNG wire#powerrail
      "Pick_Place_DB"()
      "Place_DB_7"()
   END_RUNG
   // the same network as SCL:
   "Pick_Place_DB"(ENO => #_w1);   // "Pick_Hafif"
   IF #_w1 THEN
       "Place_DB_7"();   // "Place_Hafif"
   END_IF;
END_REGION

REGION Network 8
   RUNG wire#powerrail
      "Pick_Ağır_DB"()
      "Place_Ağır_DB"()
   END_RUNG
   // the same network as SCL:
   "Pick_Ağır_DB"(ENO => #_w1);   // "Pick_Ağır"
   IF #_w1 THEN
       "Place_Ağır_DB"();   // "Place_Ağır"
   END_IF;
END_REGION

REGION Network 9
   RUNG wire#powerrail
      "Pick_Orta_DB"()
      "Place_Orta_DB"()
   END_RUNG
   // the same network as SCL:
   "Pick_Orta_DB"(ENO => #_w1);   // "Pick_Orta"
   IF #_w1 THEN
       "Place_Orta_DB"();   // "Place_Orta"
   END_IF;
END_REGION

REGION Network 10
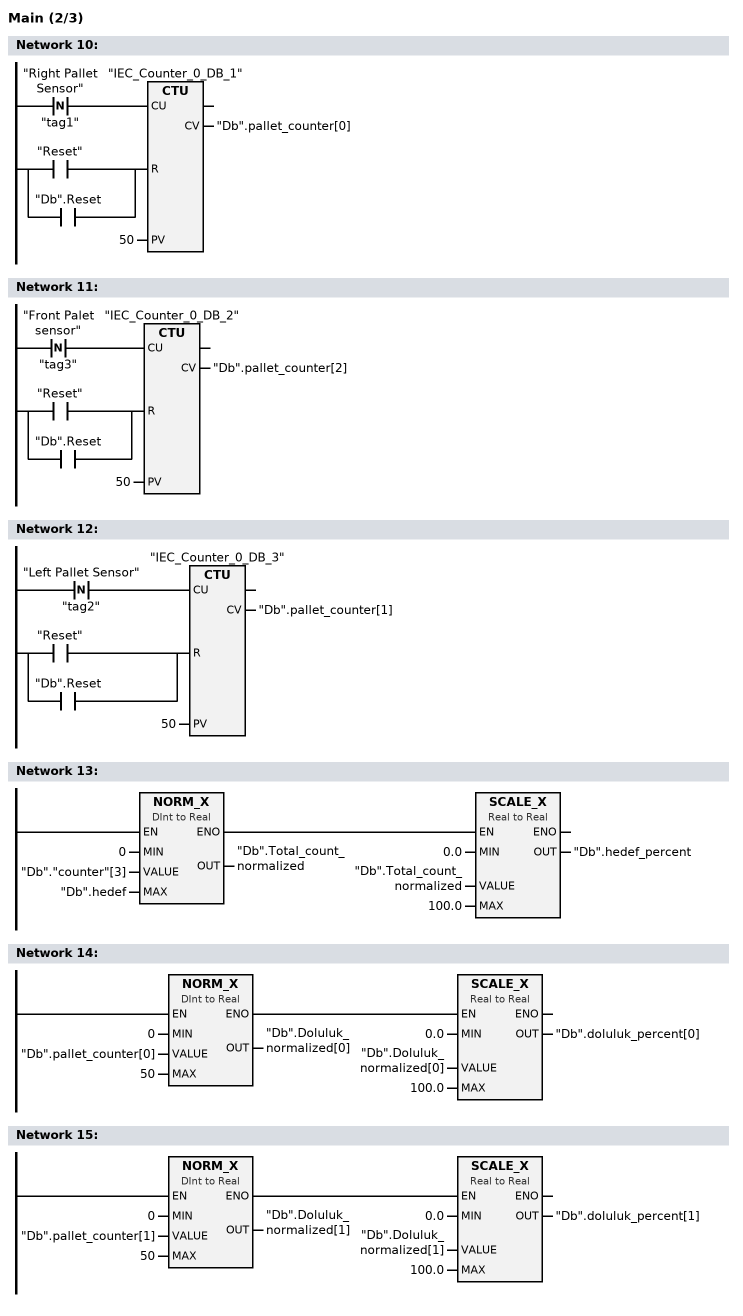
   #_w1 := NOT "Right Pallet Sensor" AND "tag1";   // falling edge of "Right Pallet Sensor"
   "tag1" := "Right Pallet Sensor";
   "IEC_Counter_0_DB_1".CTU(CU := #_w1, R := "Reset" OR "Db".Reset, PV := 50, CV => "Db".pallet_counter[0]);
END_REGION

REGION Network 11
   #_w1 := NOT "Front Palet sensor" AND "tag3";   // falling edge of "Front Palet sensor"
   "tag3" := "Front Palet sensor";
   "IEC_Counter_0_DB_2".CTU(CU := #_w1, R := "Reset" OR "Db".Reset, PV := 50, CV => "Db".pallet_counter[2]);
END_REGION

REGION Network 12
   #_w1 := NOT "Left Pallet Sensor" AND "tag2";   // falling edge of "Left Pallet Sensor"
   "tag2" := "Left Pallet Sensor";
   "IEC_Counter_0_DB_3".CTU(CU := #_w1, R := "Reset" OR "Db".Reset, PV := 50, CV => "Db".pallet_counter[1]);
END_REGION

REGION Network 13
   RUNG wire#powerrail
      { S7_Templates := "[SrcType := DInt, DestType := Real]" } Normalize(min := 0, value := "Db"."counter"[3], max := "Db".hedef, out => "Db".Total_count_normalized)
      { S7_Templates := "[SrcType := Real, DestType := Real]" } Scale(min := 0.0, value := "Db".Total_count_normalized, max := 100.0, out => "Db".hedef_percent)
   END_RUNG
   // the same network as SCL:
   "Db".Total_count_normalized := NORM_X(MIN := 0, VALUE := "Db"."counter"[3], MAX := "Db".hedef);
   "Db".hedef_percent := SCALE_X(MIN := 0.0, VALUE := "Db".Total_count_normalized, MAX := 100.0);
END_REGION

REGION Network 14
   RUNG wire#powerrail
      { S7_Templates := "[SrcType := DInt, DestType := Real]" } Normalize(min := 0, value := "Db".pallet_counter[0], max := 50, out => "Db".Doluluk_normalized[0])
      { S7_Templates := "[SrcType := Real, DestType := Real]" } Scale(min := 0.0, value := "Db".Doluluk_normalized[0], max := 100.0, out => "Db".doluluk_percent[0])
   END_RUNG
   // the same network as SCL:
   "Db".Doluluk_normalized[0] := NORM_X(MIN := 0, VALUE := "Db".pallet_counter[0], MAX := 50);
   "Db".doluluk_percent[0] := SCALE_X(MIN := 0.0, VALUE := "Db".Doluluk_normalized[0], MAX := 100.0);
END_REGION

REGION Network 15
   RUNG wire#powerrail
      { S7_Templates := "[SrcType := DInt, DestType := Real]" } Normalize(min := 0, value := "Db".pallet_counter[1], max := 50, out => "Db".Doluluk_normalized[1])
      { S7_Templates := "[SrcType := Real, DestType := Real]" } Scale(min := 0.0, value := "Db".Doluluk_normalized[1], max := 100.0, out => "Db".doluluk_percent[1])
   END_RUNG
   // the same network as SCL:
   "Db".Doluluk_normalized[1] := NORM_X(MIN := 0, VALUE := "Db".pallet_counter[1], MAX := 50);
   "Db".doluluk_percent[1] := SCALE_X(MIN := 0.0, VALUE := "Db".Doluluk_normalized[1], MAX := 100.0);
END_REGION

REGION Network 16
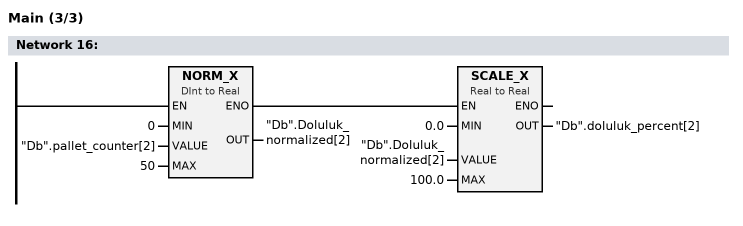
   RUNG wire#powerrail
      { S7_Templates := "[SrcType := DInt, DestType := Real]" } Normalize(min := 0, value := "Db".pallet_counter[2], max := 50, out => "Db".Doluluk_normalized[2])
      { S7_Templates := "[SrcType := Real, DestType := Real]" } Scale(min := 0.0, value := "Db".Doluluk_normalized[2], max := 100.0, out => "Db".doluluk_percent[2])
   END_RUNG
   // the same network as SCL:
   "Db".Doluluk_normalized[2] := NORM_X(MIN := 0, VALUE := "Db".pallet_counter[2], MAX := 50);
   "Db".doluluk_percent[2] := SCALE_X(MIN := 0.0, VALUE := "Db".Doluluk_normalized[2], MAX := 100.0);
END_REGION
END_ORGANIZATION_BLOCK

ORGANIZATION_BLOCK "Cyclic interrupt"   // OB30, LAD, CyclicInterrupt
{ S7_Optimized_Access := 'TRUE' }
VERSION : 0.1
   VAR_INPUT
      Initial_Call : Bool;   // Initial call of this OB
      Event_Count : Int;   // Events discarded
   END_VAR
BEGIN

REGION Network 1
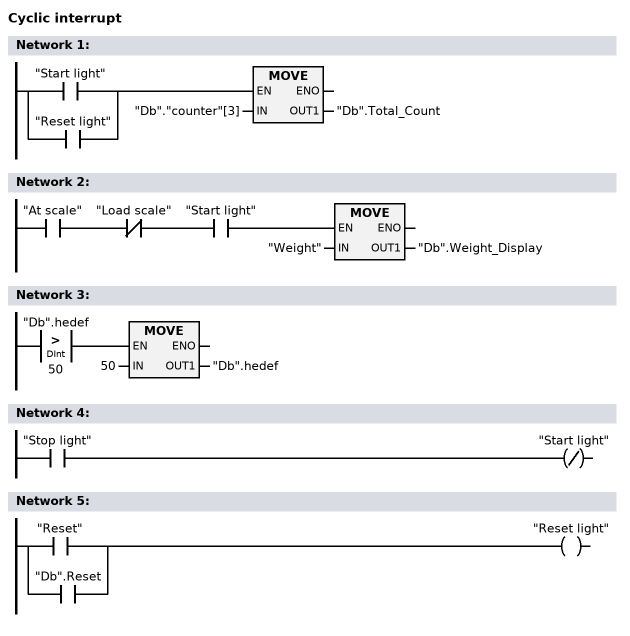
   RUNG wire#powerrail
      Contact( "Start light" )
      wire#w1
      Move(in := "Db"."counter"[3], out1 => "Db".Total_Count)
   END_RUNG
   RUNG wire#powerrail
      Contact( "Reset light" )
   END_RUNG wire#w1
   // the same network as SCL:
   IF "Start light" OR "Reset light" THEN "Db".Total_Count := "Db"."counter"[3]; END_IF;
END_REGION

REGION Network 2
   RUNG wire#powerrail
      Contact( "At scale" )
      I_Contact( "Load scale" )
      Contact( "Start light" )
      Move(in := "Weight", out1 => "Db".Weight_Display)
   END_RUNG
   // the same network as SCL:
   IF "At scale" AND NOT "Load scale" AND "Start light" THEN "Db".Weight_Display := "Weight"; END_IF;
END_REGION

REGION Network 3
   RUNG wire#powerrail
      { S7_Templates := "SrcType := DInt" } GT_Contact(in1 := "Db".hedef, in2 := 50)
      Move(in := 50, out1 => "Db".hedef)
   END_RUNG
   // the same network as SCL:
   IF "Db".hedef > 50 THEN "Db".hedef := 50; END_IF;
END_REGION

REGION Network 4
   RUNG wire#powerrail
      Contact( "Stop light" )
      I_Coil( "Start light" )
   END_RUNG
   // the same network as SCL:
   "Start light" := NOT "Stop light";
END_REGION

REGION Network 5
   RUNG wire#powerrail
      Contact( "Reset" )
      wire#w1
      Coil( "Reset light" )
   END_RUNG
   RUNG wire#powerrail
      Contact( "Db".Reset )
   END_RUNG wire#w1
   // the same network as SCL:
   "Reset light" := "Reset" OR "Db".Reset;
END_REGION
END_ORGANIZATION_BLOCK

ORGANIZATION_BLOCK "Cyclic interrupt_1"   // OB31, LAD, CyclicInterrupt
{ S7_Optimized_Access := 'TRUE' }
VERSION : 0.1
   VAR_INPUT
      Initial_Call : Bool;   // Initial call of this OB
      Event_Count : Int;   // Events discarded
   END_VAR
BEGIN

REGION Network 1
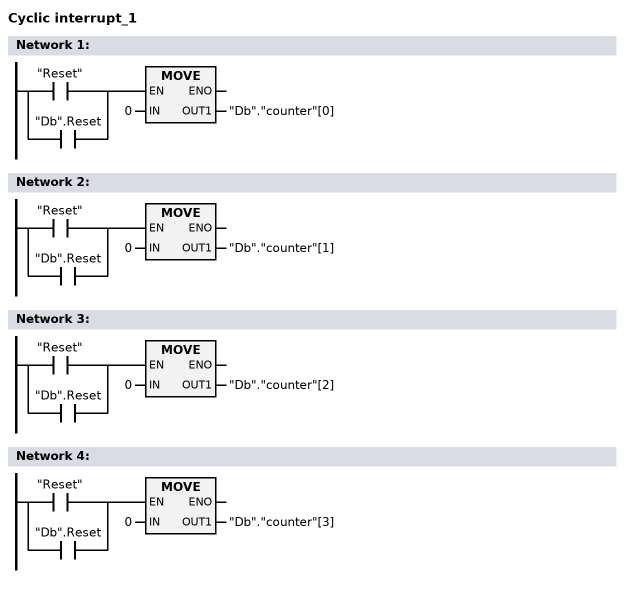
   RUNG wire#powerrail
      Contact( "Reset" )
      wire#w1
      Move(in := 0, out1 => "Db"."counter"[0])
   END_RUNG
   RUNG wire#powerrail
      Contact( "Db".Reset )
   END_RUNG wire#w1
   // the same network as SCL:
   IF "Reset" OR "Db".Reset THEN "Db"."counter"[0] := 0; END_IF;
END_REGION

REGION Network 2
   RUNG wire#powerrail
      Contact( "Reset" )
      wire#w1
      Move(in := 0, out1 => "Db"."counter"[1])
   END_RUNG
   RUNG wire#powerrail
      Contact( "Db".Reset )
   END_RUNG wire#w1
   // the same network as SCL:
   IF "Reset" OR "Db".Reset THEN "Db"."counter"[1] := 0; END_IF;
END_REGION

REGION Network 3
   RUNG wire#powerrail
      Contact( "Reset" )
      wire#w1
      Move(in := 0, out1 => "Db"."counter"[2])
   END_RUNG
   RUNG wire#powerrail
      Contact( "Db".Reset )
   END_RUNG wire#w1
   // the same network as SCL:
   IF "Reset" OR "Db".Reset THEN "Db"."counter"[2] := 0; END_IF;
END_REGION

REGION Network 4
   RUNG wire#powerrail
      Contact( "Reset" )
      wire#w1
      Move(in := 0, out1 => "Db"."counter"[3])
   END_RUNG
   RUNG wire#powerrail
      Contact( "Db".Reset )
   END_RUNG wire#w1
   // the same network as SCL:
   IF "Reset" OR "Db".Reset THEN "Db"."counter"[3] := 0; END_IF;
END_REGION
END_ORGANIZATION_BLOCK

(* ===== HMI "HMI_RT_1" =====
system functions are stored by id; their names below are inferred from use
connection "HMI_Connection_1": ETHERNET, SMART_S7_1200_OMS

HMI tags "Default tag table"
   "At scale entry" : Bool = PLC "At scale entry" AT %I0.0, 100 ms
   "At scale" : Bool = PLC "At scale" AT %I0.1, 100 ms
   "At scale exit" : Bool = PLC "At scale exit" AT %I0.2, 100 ms
   "At exit left" : Bool = PLC "At exit left" AT %I0.4, 100 ms
   "At exit front" : Bool = PLC "At exit front" AT %I0.6, 100 ms
   "At exit right" : Bool = PLC "At exit right" AT %I1.0, 100 ms
   "Reset" : Bool = PLC Reset AT %I1.2, 100 ms
   "FACTORY I/O (Running)" : Bool = PLC "FACTORY I/O (Running)" AT %I1.5, 100 ms
   "Entry conveyor" : Bool = PLC "Entry conveyor" AT %Q0.0, 100 ms
   "Load scale" : Bool = PLC "Load scale" AT %Q0.1, 100 ms
   "Right conveyor" : Bool = PLC "Right conveyor" AT %Q0.5, 100 ms
   "Reset light" : Bool = PLC "Reset light" AT %Q1.1, 100 ms
   "Weight" : Real = PLC Weight AT %ID30, 100 ms
   "Db_Weight_Value{0}" : Real = PLC "Db".Weight_Value[0], 100 ms
   "Db_Weight_Value{1}" : Real = PLC "Db".Weight_Value[1], 100 ms
   "Db_Weight_Value{2}" : Real = PLC "Db".Weight_Value[2], 100 ms
   "Db_Weight_Value{3}" : Real = PLC "Db".Weight_Value[3], 100 ms
   "Db_Weight_Value{4}" : Real = PLC "Db".Weight_Value[4], 100 ms
   "Db_hedef" : DInt = PLC "Db".hedef, 100 ms
   "Db_hedef_percent" : Real = PLC "Db".hedef_percent, 100 ms
   "Db_doluluk_percent{1}" : Real = PLC "Db".doluluk_percent[1], 100 ms
   "Db_counter{0}" : DInt = PLC "Db".counter[0], 100 ms
   "Db_pallet_counter{0}" : DInt = PLC "Db".pallet_counter[0], 100 ms
   "Db_Tartı_Hız" : Time = PLC "Db".Tartı_Hız, 100 ms
   "Db_Pick_Place_Hız" : Time = PLC "Db".Pick_Place_Hız, 100 ms
   "Db_pallet_counter{1}" : DInt = PLC "Db".pallet_counter[1], 100 ms
   "Db_counter{1}" : DInt = PLC "Db".counter[1], 100 ms
   "Db_doluluk_percent{0}" : Real = PLC "Db".doluluk_percent[0], 100 ms
   "Db_counter{2}" : DInt = PLC "Db".counter[2], 100 ms
   "Db_pallet_counter{2}" : DInt = PLC "Db".pallet_counter[2], 100 ms
   "Db_doluluk_percent{2}" : Real = PLC "Db".doluluk_percent[2], 100 ms
   "Db_Start" : Bool = PLC "Db".Start, 100 ms
   "Db_Stop" : Bool = PLC "Db".Stop, 100 ms
   "Db_Reset" : Bool = PLC "Db".Reset, 100 ms
   "Db_Weight_Display" : Real = PLC "Db".Weight_Display, 1 s
   "Db_Enable" : Bool = PLC "Db".Enable, 100 ms

text list "Tartı Ölçüm Hızı": 500 'Hızlı'; 1000 'Orta'; 1500 'Yavaş'

text list "Paletleme Hızı": 500 'Hızlı'; 1000 'Orta'; 1500 'Yavaş'

recipe "Reçete Ekranı": Hafif_Min <- "Db_Weight_Value{0}", Hafif_Max <- "Db_Weight_Value{1}", Orta_Min <- "Db_Weight_Value{2}", Orta_Max <- "Db_Weight_Value{3}", Ağır <- "Db_Weight_Value{4}", Hedef <- "Db_hedef"

Template "Template_1" 800x480
   Button "Exit" at 714,429 size 71x50; TextOff 'Exit'; PictureOff "ExitRuntime_KTP700_Basic_PN_TR"; PictureOn "ExitRuntime_KTP700_Basic_PN_TR"
      on Release: StopRuntime(0)
   Button "Log on" at 3,429 size 71x50; TextOff 'Log on'; PictureOff "Login_KTP700_Basic_PN_TR"; PictureOn "Login_KTP700_Basic_PN_TR"
      on Release: function_a2a04561()
   DateTimeField "Template_Date/time field_1" at 581,7 size 219x32
   TextField "Template_Text field_1" at 88,91 size 640x43; Text 'Akıllı Paletleme Sistemine Hoşgeldiniz!!'
   Button "HmiScreenItemData" at 81,270 size 159x47; TextOn 'Screen2'; TextOff 'Hafif Yük Hattı'; PictureOn "Navigates to Screen2 for KTP700 Basic+ PN 16.0.0.0"; PictureOff "Navigates to Screen2 for KTP700 Basic+ PN 16.0.0.0"; Authorization "Hafif_Yük_Hattı"
      on Release: ActivateScreen("Hafif Yük Hattı", 0)
   Button "HmiScreenItemData_1" at 340,271 size 160x47; TextOn 'Hafif Yük Hattı'; TextOff 'Orta Ağırlık Yük Hattı'; PictureOn "Navigates to Screen3 for KTP700 Basic+ PN 16.0.0.0"; PictureOff "Navigates to Screen3 for KTP700 Basic+ PN 16.0.0.0"; Authorization "Orta_Yük_Hattı"
      on Release: ActivateScreen("Orta_Ağırlık_Yük Hattı", 0)
   Button "HmiScreenItemData_2" at 555,271 size 159x47; TextOn 'Screen4'; TextOff 'Ağır Yük Hattı'; PictureOn "Navigates to Screen4 for KTP700 Basic+ PN 16.0.0.0"; PictureOff "Navigates to Screen4 for KTP700 Basic+ PN 16.0.0.0"; Authorization "Ağır_Yük_Hattı"
      on Release: ActivateScreen("Ağır Yük Hattı", 0)
   Button "HmiScreenItemData_4" at 81,196 size 159x47; TextOn 'Reçete'; TextOff 'Reçete'; PictureOn "Navigates to Screen2 for KTP700 Basic+ PN 16.0.0.0"; PictureOff "Navigates to Screen2 for KTP700 Basic+ PN 16.0.0.0"; Authorization "Reçete"
      on Release: ActivateScreen("Reçete", 0)
   Button "HmiScreenItemData_3" at 341,193 size 159x47; TextOn 'Tartı'; TextOff 'Tartı'; PictureOn "Navigates to Screen2 for KTP700 Basic+ PN 16.0.0.0"; PictureOff "Navigates to Screen2 for KTP700 Basic+ PN 16.0.0.0"; Authorization "Tartı"
      on Release: ActivateScreen("Tartı", 0)
   Button "HmiScreenItemData_5" at 555,193 size 159x47; TextOn 'Reçete'; TextOff 'Misafir'; PictureOn "Navigates to Screen2 for KTP700 Basic+ PN 16.0.0.0"; PictureOff "Navigates to Screen2 for KTP700 Basic+ PN 16.0.0.0"; Authorization "Misafir"
      on Release: ActivateScreen("Misafir", 0)

screen "Reçete" 800x480, template "Template_2"
   TextField "HmiScreenItemData" at 84,200 size 640x25; Text 'Screen2'
   Button "Back" at 1,1 size 159x47; TextOff 'Back'
      on Release: ActivateScreen("Root screen", 0)
   RecipeView "Recipe view_1" at 211,89 size 400x330; Authorization "Reçete"

screen "Hafif Yük Hattı" 800x480, template "Template_2"
   Button "Back" at 1,1 size 159x47; TextOff 'Back'
      on Release: ActivateScreen("Root screen", 0)
   TextField "Text field_1" at 315,53 size 180x33; Text 'Hafif Yük Hattı'
   GraphicView "Graphic view_1" at 0,303 size 486x144; Picture "Graphic_2"
   GraphicView "Graphic view_2" at 51,303 size 107x89; Picture "Graphic_7"
      HorizontalMovement <- "Db_counter{0}"
   Bar "Bar_2" at 674,169 size 80x120; MinimumValue 0; MaximumValue 100
      ProcessValue <- "Db_hedef_percent"
   TextField "Text field_3" at 562,217 size 97x23; Text 'Hedef (%):'
   Bar "Bar_3" at 465,169 size 80x120; MinimumValue 0; MaximumValue 100
      ProcessValue <- "Db_doluluk_percent{1}"
   TextField "Text field_4" at 289,217 size 153x23; Text 'Depo Doluluk(%):'
   SymbolicIOField "Symbolic I/O field_1" at 178,169 size 96x32; TextOn '1'; TextOff '0'; TextList "Paletleme Hızı"; Authorization "Paletleme Ölçüm Hızı Ayarlama"
      ProcessValue <- "Db_Pick_Place_Hız"
   TextField "Text field_5" at 16,172 size 133x23; Text 'Pick&Place Hız:'
   IOField "I/O field_1" at 179,217 size 96x32; FormatPattern s9999999999
      ProcessValue <- "Db_counter{0}"
   TextField "Text field_2" at 16,221 size 156x23; Text 'Geçen Kutu Sayısı:'
   IOField "I/O field_2" at 178,266 size 96x32; FormatPattern s9999999999
      ProcessValue <- "Db_pallet_counter{0}"
   TextField "Text field_6" at 10,266 size 161x23; Text 'Geçen Palet Sayısı:'
   GraphicView "Graphic view_9" at 702,361 size 53x60; Picture "Graphic_7"
      Visibility <- "At exit right"
   GraphicView "Graphic view_11" at 660,402 size 128x32; Picture "Graphic_18"
   GraphicView "Graphic view_8" at 622,342 size 53x60; Picture "Graphic_7"
      Visibility <- "At exit right"
   Switch "Switch_2" at 280,101 size 64x32; CaptionText 'Switch'; TextOff 'OFF'; TextOn 'ON'; Authorization "sistem başlatma"
      ProcessValue <- "Db_Start"
   Button "Button_3" at 455,101 size 96x32; TextOff 'Stop'; Authorization "sistem durdurma"
      on Click: ResetBit("Db_Start")
   Button "Button_4" at 687,101 size 96x32; TextOff 'Reset'; Authorization "sistem resetleme"
      on Release: ResetBit("Db_Reset")
      on Press: SetBit("Db_Reset")
   TextField "Text field_7" at 204,103 size 52x23; Text 'Start:'
   IOField "I/O field_3" at 674,310 size 96x32; FormatPattern 9999999
      ProcessValue <- "Db_hedef"
   TextField "Text field_8" at 563,310 size 59x23; Text 'Hedef:'
   Switch "Switch_1" at 115,103 size 64x32; CaptionText 'Switch'; TextOff 'OFF'; TextOn 'ON'; Authorization "sistem başlatma"
      ProcessValue <- "Db_Enable"
   TextField "Text field_9" at 39,105 size 66x23; Text 'Enable:'
   GraphicView "Graphic view_3" at 1,392 size 47x47; Picture "Graphic_9"
      Visibility <- "Db_counter{0}"
   GraphicView "Graphic view_4" at 1,392 size 47x47; Picture "Graphic_13"
      Visibility <- "Db_counter{0}"
   GraphicView "Graphic view_5" at 1,392 size 47x47; Picture "Graphic_14"
      Visibility <- "Db_counter{0}"
   GraphicView "Graphic view_6" at 1,392 size 47x47; Picture "Graphic_15"
      Visibility <- "Db_counter{0}"

screen "Ağır Yük Hattı" 800x480, template "Template_2"
   Button "Back" at 1,1 size 159x47; TextOff 'Back'
      on Release: ActivateScreen("Root screen", 0)
   GraphicView "Graphic view_1" at 0,303 size 486x144; Picture "Graphic_2"
   GraphicView "Graphic view_2" at 51,303 size 107x89; Picture "Graphic_7"
      HorizontalMovement <- "Db_counter{2}"
   Bar "Bar_2" at 676,172 size 80x120; MinimumValue 0; MaximumValue 100
      ProcessValue <- "Db_hedef_percent"
   TextField "Text field_3" at 564,220 size 97x23; Text 'Hedef (%):'
   Bar "Bar_3" at 467,172 size 80x120; MinimumValue 0; MaximumValue 100
      ProcessValue <- "Db_doluluk_percent{2}"
   TextField "Text field_4" at 291,220 size 153x23; Text 'Depo Doluluk(%):'
   SymbolicIOField "Symbolic I/O field_1" at 181,175 size 96x32; TextOn '1'; TextOff '0'; TextList "Paletleme Hızı"; Authorization "Paletleme Ölçüm Hızı Ayarlama"
      ProcessValue <- "Db_Pick_Place_Hız"
   TextField "Text field_5" at 23,175 size 133x23; Text 'Pick&Place Hız:'
   IOField "I/O field_1" at 181,220 size 96x32; FormatPattern s9999999999
      ProcessValue <- "Db_counter{2}"
   TextField "Text field_2" at 18,224 size 156x23; Text 'Geçen Kutu Sayısı:'
   IOField "I/O field_2" at 180,269 size 96x32; FormatPattern s9999999999
      ProcessValue <- "Db_pallet_counter{2}"
   TextField "Text field_6" at 12,269 size 161x23; Text 'Geçen Palet Sayısı:'
   TextField "Text field_1" at 315,53 size 171x33; Text 'Ağır Yük Hattı'
   GraphicView "Graphic view_9" at 675,365 size 53x60; Picture "Graphic_7"
      HorizontalMovement <- "Db_counter{1}"
      Visibility <- "At exit front"
   GraphicView "Graphic view_11" at 633,406 size 128x32; Picture "Graphic_18"
   GraphicView "Graphic view_8" at 595,346 size 53x60; Picture "Graphic_7"
      Visibility <- "At exit front"
   IOField "I/O field_3" at 676,314 size 96x32; FormatPattern 9999999
      ProcessValue <- "Db_hedef"
   TextField "Text field_8" at 564,314 size 59x23; Text 'Hedef:'
   Switch "Switch_2" at 280,101 size 64x32; CaptionText 'Switch'; TextOff 'OFF'; TextOn 'ON'; Authorization "sistem başlatma"
      ProcessValue <- "Db_Start"
   Button "Button_3" at 455,101 size 96x32; TextOff 'Stop'; Authorization "sistem durdurma"
      on Click: ResetBit("Db_Start")
   Button "Button_4" at 687,101 size 96x32; TextOff 'Reset'; Authorization "sistem resetleme"
      on Release: ResetBit("Db_Reset")
      on Press: SetBit("Db_Reset")
   TextField "Text field_7" at 204,103 size 52x23; Text 'Start:'
   Switch "Switch_1" at 115,103 size 64x32; CaptionText 'Switch'; TextOff 'OFF'; TextOn 'ON'; Authorization "sistem başlatma"
      ProcessValue <- "Db_Enable"
   TextField "Text field_9" at 39,105 size 66x23; Text 'Enable:'
   GraphicView "Graphic view_15" at 1,392 size 47x47; Picture "Graphic_9"
      Visibility <- "Db_counter{2}"
   GraphicView "Graphic view_16" at 1,392 size 47x47; Picture "Graphic_13"
      Visibility <- "Db_counter{2}"
   GraphicView "Graphic view_17" at 1,392 size 47x47; Picture "Graphic_14"
      Visibility <- "Db_counter{2}"
   GraphicView "Graphic view_18" at 1,392 size 47x47; Picture "Graphic_15"
      Visibility <- "Db_counter{2}"

screen "Tartı" 800x480, template "Template_2"
   SymbolicIOField "Symbolic I/O field_1" at 147,347 size 96x32; TextOn '1'; TextOff '0'; TextList "Tartı Ölçüm Hızı"; Authorization "Ağırlık_Ölçüm_Hızı_Ayarlama"
      ProcessValue <- "Db_Tartı_Hız"
   TextField "Text field_5" at 0,347 size 142x23; Text 'Tartı Ölçüm Hızı:'
   GraphicView "Graphic view_2" at 291,238 size 251x186; Picture "Graphic_3"
   GraphicView "Graphic view_4" at 265,157 size 102x121; Picture "Graphic_5"
      Visibility <- "At scale entry"
   GraphicView "Graphic view_1" at 367,157 size 102x121; Picture "Graphic_5"
      Visibility <- "At scale"
   GraphicView "Graphic view_3" at 469,157 size 102x121; Picture "Graphic_5"
      Visibility <- "At scale exit"
   TextField "Text field_1" at 345,55 size 143x33; Text 'Tartı Ekranı'
   IOField "I/O field_1" at 386,302 size 96x32; FormatPattern 999999999.999
      ProcessValue <- "Db_Weight_Display"
   TextField "Text field_2" at 311,305 size 65x23; Text 'Ağırlık:'
   Switch "Switch_2" at 280,101 size 64x32; CaptionText 'Switch'; TextOff 'OFF'; TextOn 'ON'; Authorization "sistem başlatma"
      ProcessValue <- "Db_Start"
   Button "Button_3" at 455,101 size 96x32; TextOff 'Stop'; Authorization "sistem durdurma"
      on Click: ResetBit("Db_Start")
   Button "Button_4" at 687,101 size 96x32; TextOff 'Reset'; Authorization "sistem resetleme"
      on Release: ResetBit("Db_Reset")
      on Press: SetBit("Db_Reset")
   TextField "Text field_7" at 204,103 size 52x23; Text 'Start:'
   Switch "Switch_1" at 115,103 size 64x32; CaptionText 'Switch'; TextOff 'OFF'; TextOn 'ON'; Authorization "sistem başlatma"
      ProcessValue <- "Db_Enable"
   TextField "Text field_9" at 39,105 size 66x23; Text 'Enable:'

screen "Orta_Ağırlık_Yük Hattı" 800x480, template "Template_2"
   GraphicView "Graphic view_1" at 0,303 size 486x144; Picture "Graphic_2"
   Bar "Bar_2" at 670,148 size 80x120; MinimumValue 0; MaximumValue 100
      ProcessValue <- "Db_hedef_percent"
   TextField "Text field_3" at 558,196 size 97x23; Text 'Hedef (%):'
   Bar "Bar_3" at 461,148 size 80x120; MinimumValue 0; MaximumValue 100
      ProcessValue <- "Db_doluluk_percent{1}"
   TextField "Text field_4" at 285,196 size 153x23; Text 'Depo Doluluk(%):'
   SymbolicIOField "Symbolic I/O field_1" at 171,148 size 96x32; TextOn '1'; TextOff '0'; TextList "Paletleme Hızı"
      ProcessValue <- "Db_Pick_Place_Hız"
   TextField "Text field_5" at 12,151 size 133x23; Text 'Pick&Place Hız:'
   IOField "I/O field_1" at 175,196 size 96x32; FormatPattern s9999999999
      ProcessValue <- "Db_counter{1}"
   TextField "Text field_2" at 12,200 size 156x23; Text 'Geçen Kutu Sayısı:'
   IOField "I/O field_2" at 174,245 size 96x32; FormatPattern s9999999999
      ProcessValue <- "Db_pallet_counter{1}"
   TextField "Text field_6" at 6,245 size 161x23; Text 'Geçen Palet Sayısı:'
   TextField "Text field_1" at 258,49 size 258x33; Text 'Orta Ağırlık Yük Hattı'
   GraphicView "Graphic view_2" at 51,303 size 107x89; Picture "Graphic_7"
      HorizontalMovement <- "Db_counter{1}"
   GraphicView "Graphic view_9" at 682,351 size 53x60; Picture "Graphic_7"
      Visibility <- "At exit left"
   GraphicView "Graphic view_11" at 640,392 size 128x32; Picture "Graphic_18"
   GraphicView "Graphic view_8" at 602,332 size 53x60; Picture "Graphic_7"
      Visibility <- "At exit left"
   IOField "I/O field_3" at 670,290 size 96x32; FormatPattern 9999999
      ProcessValue <- "Db_hedef"
   TextField "Text field_8" at 559,290 size 59x23; Text 'Hedef:'
   Switch "Switch_2" at 280,101 size 64x32; CaptionText 'Switch'; TextOff 'OFF'; TextOn 'ON'; Authorization "sistem başlatma"
      ProcessValue <- "Db_Start"
   Button "Button_3" at 455,101 size 96x32; TextOff 'Stop'; Authorization "sistem durdurma"
      on Click: ResetBit("Db_Start")
   Button "Button_4" at 687,101 size 96x32; TextOff 'Reset'; Authorization "sistem resetleme"
      on Release: ResetBit("Db_Reset")
      on Press: SetBit("Db_Reset")
   TextField "Text field_7" at 204,103 size 52x23; Text 'Start:'
   Switch "Switch_1" at 115,103 size 64x32; CaptionText 'Switch'; TextOff 'OFF'; TextOn 'ON'; Authorization "sistem başlatma"
      ProcessValue <- "Db_Enable"
   TextField "Text field_9" at 39,105 size 66x23; Text 'Enable:'
   GraphicView "Graphic view_19" at 12,391 size 47x47; Picture "Graphic_9"
      Visibility <- "Db_counter{1}"
   GraphicView "Graphic view_20" at 12,391 size 47x47; Picture "Graphic_13"
      Visibility <- "Db_counter{1}"
   GraphicView "Graphic view_21" at 12,391 size 47x47; Picture "Graphic_14"
      Visibility <- "Db_counter{1}"
   GraphicView "Graphic view_22" at 12,391 size 47x47; Picture "Graphic_15"
      Visibility <- "Db_counter{1}"

screen "Misafir" 800x480, template "Template_2"
   Button "Back" at 1,1 size 159x47; TextOn 'Back'; TextOff 'Back'
      on Release: ActivateScreen("Root screen", 0)
   Bar "Bar_2" at 131,135 size 80x120; MinimumValue 0; MaximumValue 100
      ProcessValue <- "Db_hedef_percent"
   TextField "Text field_3" at 14,135 size 97x23; Text 'Hedef (%):'
   Bar "Bar_3" at 621,304 size 80x120; MinimumValue 0; MaximumValue 100
      ProcessValue <- "Db_doluluk_percent{0}"
   TextField "Text field_4" at 536,273 size 227x23; Text 'Hafif Yük Depo Doluluk(%)'
   Bar "Bar_1" at 95,304 size 80x115; MinimumValue 0; MaximumValue 100
      ProcessValue <- "Db_doluluk_percent{1}"
   TextField "Text field_1" at 14,273 size 247x23; Text 'Orta Ağırlık Depo Doluluk(%)'
   Bar "Bar_4" at 364,304 size 80x120; MinimumValue 0; MaximumValue 100
      ProcessValue <- "Db_doluluk_percent{2}"
   TextField "Text field_2" at 285,273 size 222x23; Text 'Ağır Yük Depo Doluluk(%)'
   IOField "I/O field_1" at 701,141 size 96x32; FormatPattern 9999999
      ProcessValue <- "Db_hedef"
   TextField "Text field_5" at 533,142 size 59x23; Text 'Hedef:'
   SymbolicIOField "Symbolic I/O field_1" at 701,183 size 96x32; TextOff '0'; TextOn '1'; TextList "Tartı Ölçüm Hızı"
      ProcessValue <- "Db_Tartı_Hız"
   TextField "Text field_6" at 530,183 size 156x23; Text 'Ağırlık Ölçüm Hızı:'
   SymbolicIOField "Symbolic I/O field_2" at 701,103 size 96x32; TextOn '1'; TextOff '0'; TextList "Paletleme Hızı"
      ProcessValue <- "Db_Pick_Place_Hız"
   TextField "Text field_7" at 533,103 size 124x23; Text 'Paletleme Hızı'
   TextField "Text field_8" at 364,80 size 117x23; Text 'Misafir Ekranı'
   IOField "I/O field_2" at 701,223 size 96x32; FormatPattern 999999999.999
      ProcessValue <- "Db_Weight_Display"
   TextField "Text field_9" at 531,228 size 65x23; Text 'Ağırlık:'

Template "Template_2" 800x480
   DateTimeField "Template_Date/time field_1" at 581,7 size 219x32
   TextField "Template_Text field_1" at 185,7 size 384x43; Text 'Akıllı Paletleme Sistemi'
   Button "Exit" at 714,429 size 71x50; TextOn 'Exit'; TextOff 'Exit'; PictureOn "ExitRuntime_KTP700_Basic_PN_TR"; PictureOff "ExitRuntime_KTP700_Basic_PN_TR"
      on Release: StopRuntime(0)
   Button "Log on" at 370,429 size 71x50; TextOn 'Log on'; TextOff 'Log on'; PictureOn "Login_KTP700_Basic_PN_TR"; PictureOff "Login_KTP700_Basic_PN_TR"
      on Release: function_a2a04561()
   Button "Start screen" at 14,429 size 71x50; TextOn 'Start screen'; TextOff 'Start screen'; PictureOn "NavigateHome_KTP700_Basic_PN_TR"; PictureOff "NavigateHome_KTP700_Basic_PN_TR"
      on Release: ActivateScreen("Root screen", 0)
*)